(* PLC project Gaia V7.project, CODESYS CODESYS V3.5 SP22 Patch 2 *)
(* stored: creationDateTime 2026-11-05T09:22:17.1049023, modificationDateTime 2026-11-05T09:04:31.1849933 *)

TYPE DUT_COM_ADM100W : STRUCT
  COM_INPUT_IR : ARRAY[0..87] OF WORD;  (* [COM : Modbus RTU, input (equipment to PLC)] Input registers 0..87, 32-bit float, MSW first (ABCD) *)
  COM_INPUT_COILS : ARRAY[0..1] OF BYTE;  (* Coils 0..9 = alarms 1..10 (byte.bit) *)
  HMI_INPUT_LOCAL_REQUEST : BOOL;  (* [HMI (local PanelView) : input (to PLC)] Coil 12 | ADM100W Local Request *)
  HMI_INPUT_AUTO_REQUEST : BOOL;  (* Coil 13 | ADM100W Auto Request *)
  HMI_OUTPUT_ALARM_1_STATUS : BOOL;  (* [HMI (local PanelView) : output (from PLC)] DI 10003 | ADM100W Alarm 1 Status *)
  HMI_OUTPUT_ALARM_2_STATUS : BOOL;  (* DI 10004 | ADM100W Alarm 2 Status *)
  HMI_OUTPUT_ALARM_3_STATUS : BOOL;  (* DI 10005 | ADM100W Alarm 3 Status *)
  HMI_OUTPUT_ALARM_4_STATUS : BOOL;  (* DI 10006 | ADM100W Alarm 4 Status *)
  HMI_OUTPUT_ALARM_5_STATUS : BOOL;  (* DI 10007 | ADM100W Alarm 5 Status *)
  HMI_OUTPUT_ALARM_6_STATUS : BOOL;  (* DI 10008 | ADM100W Alarm 6 Status *)
  HMI_OUTPUT_ALARM_7_STATUS : BOOL;  (* DI 10009 | ADM100W Alarm 7 Status *)
  HMI_OUTPUT_ALARM_8_STATUS : BOOL;  (* DI 10010 | ADM100W Alarm 8 Status *)
  HMI_OUTPUT_ALARM_9_STATUS : BOOL;  (* DI 10011 | ADM100W Alarm 9 Status *)
  HMI_OUTPUT_ALARM_10_STATUS : BOOL;  (* DI 10012 | ADM100W Alarm 10 Status *)
  HMI_OUTPUT_LOCAL_ACTIVE : BOOL;  (* DI 10018 | ADM100W Local Active *)
  HMI_OUTPUT_FREQUENCY : DUT_Union_Real_Word;  (* IR 1-2 | ADM100W Frequency | Hz *)
  HMI_OUTPUT_L1_L2_VOLTAGE : DUT_Union_Real_Word;  (* IR 3-4 | ADM100W L1-L2 Voltage | V *)
  HMI_OUTPUT_L1_N_VOLTAGE : DUT_Union_Real_Word;  (* IR 5-6 | ADM100W L1-N Voltage | V *)
  HMI_OUTPUT_L1_CURRENT : DUT_Union_Real_Word;  (* IR 7-8 | ADM100W L1 Current | A *)
  HMI_OUTPUT_L1_ACTIVE_POWER : DUT_Union_Real_Word;  (* IR 9-10 | ADM100W L1 Active Power *)
  HMI_OUTPUT_L1_APPARENT_POWER : DUT_Union_Real_Word;  (* IR 11-12 | ADM100W L1 Apparent Power *)
  HMI_OUTPUT_L1_REACTIVE_POWER : DUT_Union_Real_Word;  (* IR 13-14 | ADM100W L1 Reactive Power *)
  HMI_OUTPUT_L1_CURRENT_PHASE_ANGLE : DUT_Union_Real_Word;  (* IR 15-16 | ADM100W L1 Current Phase Angle | deg *)
  HMI_OUTPUT_L1_POWER_FACTOR : DUT_Union_Real_Word;  (* IR 17-18 | ADM100W L1 Power Factor *)
  HMI_OUTPUT_L1_VOLTAGE_THD : DUT_Union_Real_Word;  (* IR 19-20 | ADM100W L1 Voltage THD | % *)
  HMI_OUTPUT_L1_CURRENT_THD : DUT_Union_Real_Word;  (* IR 21-22 | ADM100W L1 Current THD | % *)
  HMI_OUTPUT_L1_MAX_LOAD : DUT_Union_Real_Word;  (* IR 23-24 | ADM100W L1 Max Load *)
  HMI_OUTPUT_L1_L2_VOLTAGE_PHASE_ANGLE : DUT_Union_Real_Word;  (* IR 25-26 | ADM100W L1-L2 Voltage Phase Angle | deg *)
  HMI_OUTPUT_L2_L3_VOLTAGE : DUT_Union_Real_Word;  (* IR 27-28 | ADM100W L2-L3 Voltage | V *)
  HMI_OUTPUT_L2_N_VOLTAGE : DUT_Union_Real_Word;  (* IR 29-30 | ADM100W L2-N Voltage | V *)
  HMI_OUTPUT_L2_CURRENT : DUT_Union_Real_Word;  (* IR 31-32 | ADM100W L2 Current | A *)
  HMI_OUTPUT_L2_ACTIVE_POWER : DUT_Union_Real_Word;  (* IR 33-34 | ADM100W L2 Active Power *)
  HMI_OUTPUT_L2_APPARENT_POWER : DUT_Union_Real_Word;  (* IR 35-36 | ADM100W L2 Apparent Power *)
  HMI_OUTPUT_L2_REACTIVE_POWER : DUT_Union_Real_Word;  (* IR 37-38 | ADM100W L2 Reactive Power *)
  HMI_OUTPUT_L2_CURRENT_PHASE_ANGLE : DUT_Union_Real_Word;  (* IR 39-40 | ADM100W L2 Current Phase Angle | deg *)
  HMI_OUTPUT_L2_POWER_FACTOR : DUT_Union_Real_Word;  (* IR 41-42 | ADM100W L2 Power Factor *)
  HMI_OUTPUT_L2_VOLTAGE_THD : DUT_Union_Real_Word;  (* IR 43-44 | ADM100W L2 Voltage THD | % *)
  HMI_OUTPUT_L2_CURRENT_THD : DUT_Union_Real_Word;  (* IR 45-46 | ADM100W L2 Current THD | % *)
  HMI_OUTPUT_L2_MAX_LOAD : DUT_Union_Real_Word;  (* IR 47-48 | ADM100W L2 Max Load *)
  HMI_OUTPUT_L1_L3_VOLTAGE_PHASE_ANGLE : DUT_Union_Real_Word;  (* IR 49-50 | ADM100W L1-L3 Voltage Phase Angle | deg *)
  HMI_OUTPUT_L3_L1_VOLTAGE : DUT_Union_Real_Word;  (* IR 51-52 | ADM100W L3-L1 Voltage | V *)
  HMI_OUTPUT_L3_N_VOLTAGE : DUT_Union_Real_Word;  (* IR 53-54 | ADM100W L3-N Voltage | V *)
  HMI_OUTPUT_L3_CURRENT : DUT_Union_Real_Word;  (* IR 55-56 | ADM100W L3 Current | A *)
  HMI_OUTPUT_L3_ACTIVE_POWER : DUT_Union_Real_Word;  (* IR 57-58 | ADM100W L3 Active Power *)
  HMI_OUTPUT_L3_APPARENT_POWER : DUT_Union_Real_Word;  (* IR 59-60 | ADM100W L3 Apparent Power *)
  HMI_OUTPUT_L3_REACTIVE_POWER : DUT_Union_Real_Word;  (* IR 61-62 | ADM100W L3 Reactive Power *)
  HMI_OUTPUT_L3_CURRENT_PHASE_ANGLE : DUT_Union_Real_Word;  (* IR 63-64 | ADM100W L3 Current Phase Angle | deg *)
  HMI_OUTPUT_L3_POWER_FACTOR : DUT_Union_Real_Word;  (* IR 65-66 | ADM100W L3 Power Factor *)
  HMI_OUTPUT_L3_VOLTAGE_THD : DUT_Union_Real_Word;  (* IR 67-68 | ADM100W L3 Voltage THD | % *)
  HMI_OUTPUT_L3_CURRENT_THD : DUT_Union_Real_Word;  (* IR 69-70 | ADM100W L3 Current THD | % *)
  HMI_OUTPUT_L3_MAX_LOAD : DUT_Union_Real_Word;  (* IR 71-72 | ADM100W L3 Max Load *)
  HMI_OUTPUT_INTERNAL_TEMPERATURE : DUT_Union_Real_Word;  (* IR 73-74 | ADM100W Internal Temperature *)
  HMI_OUTPUT_ACTIVE_ENERGY : DUT_Union_Real_Word;  (* IR 75-76 | ADM100W Active Energy *)
  HMI_OUTPUT_APPARENT_ENERGY : DUT_Union_Real_Word;  (* IR 77-78 | ADM100W Apparent Energy *)
  HMI_OUTPUT_REACTIVE_ENERGY : DUT_Union_Real_Word;  (* IR 79-80 | ADM100W Reactive Energy *)
  HMI_OUTPUT_TOTAL_ACTIVE_POWER : DUT_Union_Real_Word;  (* IR 81-82 | ADM100W Total Active Power *)
  HMI_OUTPUT_TOTAL_APPARENT_POWER : DUT_Union_Real_Word;  (* IR 83-84 | ADM100W Total Apparent Power *)
  HMI_OUTPUT_TOTAL_REACTIVE_POWER : DUT_Union_Real_Word;  (* IR 85-86 | ADM100W Total Reactive Power *)
  HMI_OUTPUT_ALL_PHASE_POWER_FACTOR : DUT_Union_Real_Word;  (* IR 87-88 | ADM100W All Phase Power Factor *)
END_STRUCT;
END_TYPE

TYPE DUT_COM_DIP1500 : STRUCT
  COM_INPUT_IR : ARRAY[0..4] OF WORD;  (* [COM : Modbus RTU, input (equipment to PLC)] Input registers 0x3001..0x3005 *)
  COM_INPUT_HR_COUNTERS : ARRAY[0..3] OF WORD;  (* Holding registers 0x4007..0x400A (read) *)
  COM_OUTPUT_COILS : ARRAY[0..3] OF BOOL;  (* [COM : Modbus RTU, output (PLC to equipment)] Coils 0x0001..0x0004 *)
  COM_OUTPUT_HR_CMD : ARRAY[0..5] OF WORD;  (* Holding registers 0x4001..0x4006 (write) *)
  COM_OUTPUT_HR_CONFIG : ARRAY[0..6] OF WORD;  (* Holding registers 0x400B..0x4011 (write) *)
  COM_OUTPUT_CMD_TRIGGER : BOOL;  (* Rising edge trigger of the command write channel(s), mapped in the Modbus slave I/O mapping *)
  COM_OUTPUT_CONFIG_TRIGGER : BOOL;  (* Rising edge trigger of the configuration write channel, mapped in the Modbus slave I/O mapping *)
  HMI_INPUT_MOTOR_START_STOP : BOOL;  (* [HMI (local PanelView) : input (to PLC)] Coil 3 | DIP1500 Motor Start Stop *)
  HMI_INPUT_MOTOR_DIRECTION : BOOL;  (* Coil 4 | DIP1500 Motor Direction *)
  HMI_INPUT_FLASH_SAVE : BOOL;  (* Coil 5 | DIP1500 Flash Save *)
  HMI_INPUT_OPERATION_MODE : BOOL;  (* Coil 6 | DIP1500 Operation Mode *)
  HMI_INPUT_PARAM_WRITE_ENABLE : BOOL;  (* Coil 7 | DIP1500 Parameter Write Enable *)
  HMI_INPUT_LOCAL_REQUEST : BOOL;  (* Coil 10 | DIP1500 Local Request *)
  HMI_INPUT_AUTO_REQUEST : BOOL;  (* Coil 11 | DIP1500 Auto Request *)
  HMI_INPUT_FOOT_SWITCH_INPUT_MODE : WORD;  (* HR 9 | DIP1500 Foot Switch Input Mode *)
  HMI_INPUT_LIQUID_LEVEL_INPUT_MODE : WORD;  (* HR 10 | DIP1500 Liquid Level Input Mode *)
  HMI_INPUT_STATE_OUTPUT_MODE : WORD;  (* HR 11 | DIP1500 State Output Mode *)
  HMI_INPUT_COMMUNICATION_ADDRESS : WORD;  (* HR 12 | DIP1500 Communication Address *)
  HMI_INPUT_BAUD_RATE_INDEX : WORD;  (* HR 13 | DIP1500 Baud Rate Index | index *)
  HMI_INPUT_MOTOR_SPEED : DUT_Union_Real_Word;  (* HR 1-2 | DIP1500 Motor Speed | rpm *)
  HMI_INPUT_MAX_MOTOR_SPEED : DUT_Union_Real_Word;  (* HR 3-4 | DIP1500 Max Motor Speed | rpm *)
  HMI_INPUT_RUN_TIME_OR_VOLUME_SETPOINT : DUT_Union_Real_Word;  (* HR 5-6 | DIP1500 Run Time Or Volume Setpoint | ms (time mode) / ml (volume mode) *)
  HMI_INPUT_FLOW_RATE_OR_SPEED_CALIBRATION_COEFFICIENT : DUT_Union_Real_Word;  (* HR 7-8 | DIP1500 Flow Rate Or Speed Calibration Coefficient | ml/min or rpm *)
  HMI_OUTPUT_LOCAL_ACTIVE : BOOL;  (* [HMI (local PanelView) : output (from PLC)] DI 10016 | DIP1500 Local Active *)
  HMI_OUTPUT_FIRMWARE_VERSION : WORD;  (* IR 91 | DIP1500 Firmware Version | 3+5+8 bits (major+minor+revision) *)
  HMI_OUTPUT_HARDWARE_VERSION : WORD;  (* IR 92 | DIP1500 Hardware Version | 3+5+8 bits (major+minor+revision) *)
  HMI_OUTPUT_TEMPERATURE : WORD;  (* IR 93 | DIP1500 Temperature | degC | (raw - 500) / 10 *)
  HMI_OUTPUT_FLOAT_LEVEL_ALARM : WORD;  (* IR 94 | DIP1500 Float Level Alarm *)
  HMI_OUTPUT_DIGITAL_OUTPUT_VALUE : WORD;  (* IR 95 | DIP1500 Digital Output Value *)
  HMI_OUTPUT_REAL_TIME_RUN_TIME_OR_VOLUME : DUT_Union_Real_Word;  (* IR 96-97 | DIP1500 Real-Time Run Time Or Volume | ms (time mode) / ml (volume mode) *)
  HMI_OUTPUT_ACCUMULATED_RUN_TIME_OR_VOLUME : DUT_Union_Real_Word;  (* IR 98-99 | DIP1500 Accumulated Run Time Or Volume | ms (time mode) / ml (volume mode) *)
END_STRUCT;
END_TYPE

TYPE DUT_COM_DOSENSOR : STRUCT
  HMI_INPUT_CALIBRATION_HIGH : BOOL;  (* [HMI (local PanelView) : input (to PLC)] Coil 1 | DO Calibration High *)
  HMI_INPUT_CALIBRATION_LOW : BOOL;  (* Coil 2 | DO Calibration Low *)
  HMI_INPUT_LOCAL_REQUEST : BOOL;  (* Coil 8 | DO Sensor Local Request *)
  HMI_INPUT_AUTO_REQUEST : BOOL;  (* Coil 9 | DO Sensor Auto Request *)
  HMI_OUTPUT_FAULT : BOOL;  (* [HMI (local PanelView) : output (from PLC)] DI 10001 | Do sensor fault *)
  HMI_OUTPUT_CALIBRATION_DONE : BOOL;  (* DI 10002 | Do sensor calibration done *)
  HMI_OUTPUT_LOCAL_ACTIVE : BOOL;  (* DI 10014 | DO Sensor Local Active *)
  HMI_OUTPUT_SIGNAL : DUT_Union_Real_Word;  (* IR 89-90 | DO Sensor Signal *)
END_STRUCT;
END_TYPE

TYPE DUT_COM_UPI_LOCAL_HMI : STRUCT
  HMI_INPUT_LOCAL_REQUEST : BOOL;  (* [HMI (local PanelView) : input (to PLC)] Coil 14 | Global Local HMI Request *)
  HMI_INPUT_AUTO_REQUEST : BOOL;  (* Coil 15 | Global Auto HMI Request *)
  HMI_OUTPUT_LOCAL_ACTIVE : BOOL;  (* [HMI (local PanelView) : output (from PLC)] DI 10020 | Global Local HMI Active *)
END_STRUCT;
END_TYPE

TYPE DUT_EXC_ADM100W : STRUCT
  EXC_OUTPUT_FREQUENCY : REAL;  (* [EXC : to other equipment] Hz *)
  EXC_OUTPUT_L1_N_VOLTAGE : REAL;  (* V *)
  EXC_OUTPUT_L1_CURRENT : REAL;  (* A *)
  EXC_OUTPUT_L1_ACTIVE_POWER : REAL;  (* W *)
  EXC_OUTPUT_L1_APPARENT_POWER : REAL;  (* VA *)
  EXC_OUTPUT_L1_REACTIVE_POWER : REAL;  (* VAr *)
  EXC_OUTPUT_L1_POWER_FACTOR : REAL;  (* - *)
  EXC_OUTPUT_L1_VOLTAGE_THD : REAL;  (* % *)
  EXC_OUTPUT_L1_CURRENT_THD : REAL;  (* % *)
  EXC_OUTPUT_L1_MAX_LOAD : REAL;  (* % of 60 A *)
  EXC_OUTPUT_INTERNAL_TEMPERATURE : REAL;  (* degC *)
  EXC_OUTPUT_ACTIVE_ENERGY : REAL;  (* kWh *)
  EXC_OUTPUT_DATA_VALID : BOOL;  (* FALSE = values not usable. Not managed yet (no Modbus diagnostic) *)
  UPI_INPUT_GLOBAL_LOCAL_HMI : BOOL;  (* [UPI : functional units to equipment] From UPI_LOCAL_HMI : global HMI local active *)
END_STRUCT;
END_TYPE

TYPE DUT_EXC_DIP1500 : STRUCT
  UPI_INPUT_GLOBAL_LOCAL_HMI : BOOL;  (* [UPI : functional units to equipment] From UPI_LOCAL_HMI : global HMI local active *)
  UPI_INPUT_RUN : BOOL;  (* [UPI : commands used in auto mode] Auto mode command : run *)
  UPI_INPUT_CLOCKWISE : BOOL;  (* Auto mode command : 1 clockwise *)
  UPI_INPUT_VOLUME_MODE : BOOL;  (* Auto mode command : 0 time mode, 1 volume mode *)
  UPI_INPUT_SPEED : REAL;  (* Auto mode command : speed, rpm *)
  UPI_INPUT_RUN_SETPOINT : REAL;  (* Auto mode command : ms (time mode) or ml (volume mode), 0 = continuous *)
END_STRUCT;
END_TYPE

TYPE DUT_EXC_DOSENSOR : STRUCT
  EXC_OUTPUT_SIGNAL : REAL;  (* [EXC : to other equipment] Dissolved oxygen measure *)
  UPI_INPUT_GLOBAL_LOCAL_HMI : BOOL;  (* [UPI : functional units to equipment] From UPI_LOCAL_HMI : global HMI local active *)
END_STRUCT;
END_TYPE

TYPE DUT_EXC_UPI_LOCAL_HMI : STRUCT
  UPI_OUTPUT_LOCAL_ACTIVE : BOOL;  (* [UPI : to equipment] Global HMI local active *)
END_STRUCT;
END_TYPE

TYPE DUT_INT_ADM100W : STRUCT
  HMI_LOCAL_REQUEST : BOOL;  (* [Control mode] From HMI : local request (pulse or maintained) *)
  HMI_AUTO_REQUEST : BOOL;  (* From HMI : auto request, releases the individual HMI local *)
  GLOBAL_LOCAL_HMI : BOOL;  (* From UPI_LOCAL_HMI : global HMI local active *)
  LOCAL_HMI_INDIVIDUAL : BOOL;  (* Memory : individual HMI local, set by local request, reset by auto request *)
  LOCAL_HMI : BOOL;  (* Result : equipment in HMI local (individual or global) *)
  AUTO : BOOL;  (* Result : no local mode, commands come from the functional units (UPI) *)
  ALARM_1 : BOOL;  (* [Alarms] Alarm 1 status *)
  ALARM_2 : BOOL;  (* Alarm 2 status *)
  ALARM_3 : BOOL;  (* Alarm 3 status *)
  ALARM_4 : BOOL;  (* Alarm 4 status *)
  ALARM_5 : BOOL;  (* Alarm 5 status *)
  ALARM_6 : BOOL;  (* Alarm 6 status *)
  ALARM_7 : BOOL;  (* Alarm 7 status *)
  ALARM_8 : BOOL;  (* Alarm 8 status *)
  ALARM_9 : BOOL;  (* Alarm 9 status *)
  ALARM_10 : BOOL;  (* Alarm 10 status *)
  FREQUENCY : REAL;  (* [Measures] Frequency | Hz *)
  L1_L2_VOLTAGE : REAL;  (* L1-L2 Voltage | V *)
  L1_N_VOLTAGE : REAL;  (* L1-N Voltage | V *)
  L1_CURRENT : REAL;  (* L1 Current | A *)
  L1_ACTIVE_POWER : REAL;  (* L1 Active Power | W *)
  L1_APPARENT_POWER : REAL;  (* L1 Apparent Power | VA *)
  L1_REACTIVE_POWER : REAL;  (* L1 Reactive Power | W *)
  L1_CURRENT_PHASE_ANGLE : REAL;  (* L1 Current Phase Angle | deg *)
  L1_POWER_FACTOR : REAL;  (* L1 Power Factor | - *)
  L1_VOLTAGE_THD : REAL;  (* L1 Voltage THD | % *)
  L1_CURRENT_THD : REAL;  (* L1 Current THD | % *)
  L1_MAX_LOAD : REAL;  (* L1 Max Load | % of 60 A *)
  L1_L2_VOLTAGE_PHASE_ANGLE : REAL;  (* L1-L2 Voltage Phase Angle | deg *)
  L2_L3_VOLTAGE : REAL;  (* L2-L3 Voltage | V *)
  L2_N_VOLTAGE : REAL;  (* L2-N Voltage | V *)
  L2_CURRENT : REAL;  (* L2 Current | A *)
  L2_ACTIVE_POWER : REAL;  (* L2 Active Power | W *)
  L2_APPARENT_POWER : REAL;  (* L2 Apparent Power | VA *)
  L2_REACTIVE_POWER : REAL;  (* L2 Reactive Power | W *)
  L2_CURRENT_PHASE_ANGLE : REAL;  (* L2 Current Phase Angle | deg *)
  L2_POWER_FACTOR : REAL;  (* L2 Power Factor | - *)
  L2_VOLTAGE_THD : REAL;  (* L2 Voltage THD | % *)
  L2_CURRENT_THD : REAL;  (* L2 Current THD | % *)
  L2_MAX_LOAD : REAL;  (* L2 Max Load | % of 60 A *)
  L1_L3_VOLTAGE_PHASE_ANGLE : REAL;  (* L1-L3 Voltage Phase Angle | deg *)
  L3_L1_VOLTAGE : REAL;  (* L3-L1 Voltage | V *)
  L3_N_VOLTAGE : REAL;  (* L3-N Voltage | V *)
  L3_CURRENT : REAL;  (* L3 Current | A *)
  L3_ACTIVE_POWER : REAL;  (* L3 Active Power | W *)
  L3_APPARENT_POWER : REAL;  (* L3 Apparent Power | VA *)
  L3_REACTIVE_POWER : REAL;  (* L3 Reactive Power | W *)
  L3_CURRENT_PHASE_ANGLE : REAL;  (* L3 Current Phase Angle | deg *)
  L3_POWER_FACTOR : REAL;  (* L3 Power Factor | - *)
  L3_VOLTAGE_THD : REAL;  (* L3 Voltage THD | % *)
  L3_CURRENT_THD : REAL;  (* L3 Current THD | % *)
  L3_MAX_LOAD : REAL;  (* L3 Max Load | % of 60 A *)
  INTERNAL_TEMPERATURE : REAL;  (* Internal Temperature | degC *)
  ACTIVE_ENERGY : REAL;  (* Active Energy | kWh *)
  APPARENT_ENERGY : REAL;  (* Apparent Energy | per ADM100W config *)
  REACTIVE_ENERGY : REAL;  (* Reactive Energy | kWh *)
  TOTAL_ACTIVE_POWER : REAL;  (* Total Active Power | W *)
  TOTAL_APPARENT_POWER : REAL;  (* Total Apparent Power | VA *)
  TOTAL_REACTIVE_POWER : REAL;  (* Total Reactive Power | W *)
  ALL_PHASE_POWER_FACTOR : REAL;  (* All Phase Power Factor | - *)
END_STRUCT;
END_TYPE

TYPE DUT_INT_DIP1500 : STRUCT
  HMI_LOCAL_REQUEST : BOOL;  (* [Control mode] From HMI : local request (pulse or maintained) *)
  HMI_AUTO_REQUEST : BOOL;  (* From HMI : auto request, releases the individual HMI local *)
  GLOBAL_LOCAL_HMI : BOOL;  (* From UPI_LOCAL_HMI : global HMI local active *)
  LOCAL_HMI_INDIVIDUAL : BOOL;  (* Memory : individual HMI local, set by local request, reset by auto request *)
  LOCAL_HMI : BOOL;  (* Result : equipment in HMI local (individual or global) *)
  AUTO : BOOL;  (* Result : no local mode, commands come from the functional units (UPI) *)
  CMD_RUN : BOOL;  (* [Commands (to pump), from the active source] 0 stop, 1 start *)
  CMD_CLOCKWISE : BOOL;  (* 0 counterclockwise, 1 clockwise *)
  CMD_SAVE_FLASH : BOOL;  (* 1 s pulse to coil 0x0003, saves pump parameters to flash *)
  CMD_VOLUME_MODE : BOOL;  (* 0 time mode, 1 volume mode *)
  CMD_SPEED : REAL;  (* rpm *)
  CMD_MAX_SPEED : REAL;  (* rpm *)
  CMD_RUN_SETPOINT : REAL;  (* ms (time mode) or ml (volume mode), 0 = continuous *)
  CMD_CALIB_COEF : REAL;  (* ml/min or rpm *)
  CMD_FOOT_MODE : WORD;  (* Foot switch input mode *)
  CMD_LEVEL_MODE : WORD;  (* Liquid level input mode *)
  CMD_STATE_OUT_MODE : WORD;  (* State output mode *)
  CMD_ADDRESS : WORD;  (* Modbus address *)
  CMD_BAUD_INDEX : WORD;  (* 0=1200 .. 3=9600 .. 7=115200 *)
  PARAM_WRITE_ENABLE : BOOL;  (* [Parameter writing] 1 = write configuration to the pump, 0 = stop writing *)
  FLASH_SAVE_REQUEST : BOOL;  (* Flash save request (rising edge used) *)
  PARAM_VALID : BOOL;  (* Address 1..31, baud index 0..7, max speed > 0, calibration coefficient > 0 *)
  PULSE_500MS : BOOL;  (* [Write triggers] Square wave, 500 ms period, source of the trigger edges *)
  CMD_CHANGED : BOOL;  (* A command value changed this cycle *)
  CMD_WINDOW : BOOL;  (* Command write window, 3 s after the last change *)
  CMD_TRIGGER : BOOL;  (* Command channel trigger *)
  CONFIG_TRIGGER : BOOL;  (* Configuration channel trigger *)
  PREV_RUN : BOOL;  (* [Previous command values] Previous values for change detection *)
  PREV_CLOCKWISE : BOOL;
  PREV_VOLUME_MODE : BOOL;
  PREV_SAVE_FLASH : BOOL;
  PREV_SPEED : REAL;
  PREV_MAX_SPEED : REAL;
  PREV_RUN_SETPOINT : REAL;
  FBK_FIRMWARE_VERSION : WORD;  (* [Feedback (from pump)] 3+5+8 bits (major+minor+revision) *)
  FBK_HARDWARE_VERSION : WORD;  (* 3+5+8 bits (major+sub+reserved) *)
  FBK_TEMPERATURE : WORD;  (* (raw - 500) / 10 = degC, 65535 = not connected *)
  FBK_LEVEL_ALARM : WORD;  (* 0 no alarm, 1 alarm, 65535 = not connected *)
  FBK_DIGITAL_OUTPUT : WORD;  (* Digital output value *)
  FBK_RUN_ACTUAL : REAL;  (* Current run, ms (time mode) or ml (volume mode) *)
  FBK_RUN_TOTAL : REAL;  (* Accumulated run, ms (time mode) or ml (volume mode) *)
  UDINT_TEMP : UDINT;  (* [Work] Work variable, time mode conversion *)
  SRC_MAX_MOTOR_SPEED : REAL;  (* [Parameter source] Value typed in the active local supervision *)
  SRC_CALIBRATION_COEFFICIENT : REAL;
  SRC_FOOT_SWITCH_INPUT_MODE : WORD;
  SRC_LIQUID_LEVEL_INPUT_MODE : WORD;
  SRC_STATE_OUTPUT_MODE : WORD;
  SRC_COMMUNICATION_ADDRESS : WORD;
  SRC_BAUD_RATE_INDEX : WORD;
  PREV_SRC_MAX_MOTOR_SPEED : REAL;  (* [Parameter change detection] Previous source values *)
  PREV_SRC_CALIBRATION_COEFFICIENT : REAL;
  PREV_SRC_FOOT_SWITCH_INPUT_MODE : WORD;
  PREV_SRC_LIQUID_LEVEL_INPUT_MODE : WORD;
  PREV_SRC_STATE_OUTPUT_MODE : WORD;
  PREV_SRC_COMMUNICATION_ADDRESS : WORD;
  PREV_SRC_BAUD_RATE_INDEX : WORD;
  PREV_LOCAL_HMI : BOOL;
  SOURCE_CHANGED : BOOL;  (* The active local source changed this cycle : no parameter is taken *)
END_STRUCT;
END_TYPE

TYPE DUT_INT_DOSENSOR : STRUCT
  HMI_LOCAL_REQUEST : BOOL;  (* [Control mode] From HMI : local request (pulse or maintained) *)
  HMI_AUTO_REQUEST : BOOL;  (* From HMI : auto request, releases the individual HMI local *)
  GLOBAL_LOCAL_HMI : BOOL;  (* From UPI_LOCAL_HMI : global HMI local active *)
  LOCAL_HMI_INDIVIDUAL : BOOL;  (* Memory : individual HMI local, set by local request, reset by auto request *)
  LOCAL_HMI : BOOL;  (* Result : equipment in HMI local (individual or global) *)
  AUTO : BOOL;  (* Result : no local mode, commands come from the functional units (UPI) *)
  SIGNAL_RAW : DWORD;  (* [Inputs] Raw analog input *)
  FAULT : BOOL;  (* Sensor fault (digital input) *)
  CALIB_HIGH_REQUEST : BOOL;  (* High calibration request from the active source *)
  CALIB_LOW_REQUEST : BOOL;  (* Low calibration request from the active source *)
  SIGNAL : REAL;  (* [Results] Scaled measure *)
  CALIB_HIGH : BOOL;  (* High calibration pulse to sensor (1 s) *)
  CALIB_LOW : BOOL;  (* Low calibration pulse to sensor (1 s) *)
  CALIB_DONE : BOOL;  (* Calibration done message (5 s) *)
END_STRUCT;
END_TYPE

TYPE DUT_INT_UPI_LOCAL_HMI : STRUCT
  LOCAL_REQUEST : BOOL;  (* Local request (pulse or maintained) *)
  AUTO_REQUEST : BOOL;  (* Auto request, releases the global local *)
  LOCAL_ACTIVE : BOOL;  (* Memory : global local active *)
END_STRUCT;
END_TYPE

TYPE DUT_IO_ADM100W : STRUCT
  SPARE : BOOL;  (* Placeholder, structure not used yet *)
END_STRUCT;
END_TYPE

TYPE DUT_IO_DIP1500 : STRUCT
  SPARE : BOOL;  (* Placeholder, structure not used yet *)
END_STRUCT;
END_TYPE

TYPE DUT_IO_DOSENSOR : STRUCT
  INPUT_SIGNAL : DWORD;  (* [INPUT (field to PLC)] Analog input, raw value *)
  INPUT_SENSOR_FAULT : BOOL;  (* Digital input, sensor fault *)
  OUTPUT_CALIBRATION_HIGH : BOOL;  (* [OUTPUT (PLC to field)] Digital output, high calibration *)
  OUTPUT_CALIBRATION_LOW : BOOL;  (* Digital output, low calibration *)
END_STRUCT;
END_TYPE

TYPE DUT_PA_ADM100W : STRUCT
  SPARE : BOOL;  (* Placeholder, structure not used yet *)
END_STRUCT;
END_TYPE

TYPE DUT_PA_DIP1500 : STRUCT
  MAX_MOTOR_SPEED : REAL := 350;  (* [Pump configuration, default value = declaration value, kept in GVL_PA (persistent)] rpm. Max motor speed (pump register 0x4003) *)
  CALIBRATION_COEFFICIENT : REAL := 100;  (* ml/min or rpm. Flow / speed calibration coefficient (0x400B) *)
  FOOT_SWITCH_INPUT_MODE : WORD := 0;  (* Foot switch input mode (0x400D) *)
  LIQUID_LEVEL_INPUT_MODE : WORD := 100;  (* Liquid level input mode (0x400E) *)
  STATE_OUTPUT_MODE : WORD := 7;  (* State output mode (0x400F) *)
  COMMUNICATION_ADDRESS : WORD := 11;  (* Pump Modbus address, 1..31 (0x4010) *)
  BAUD_RATE_INDEX : WORD := 3;  (* 0=1200 .. 3=9600 .. 7=115200 (0x4011) *)
END_STRUCT;
END_TYPE

TYPE DUT_PA_DOSENSOR : STRUCT
  SPARE : BOOL;  (* Placeholder, structure not used yet *)
END_STRUCT;
END_TYPE

TYPE DUT_Union_Real_Word : UNION
  Real_value : REAL;
  Word_value : ARRAY[0..1] OF WORD;
END_UNION;
END_TYPE

FUNCTION_BLOCK FB_INST_ADM100W
  VAR_IN_OUT
    PA : DUT_PA_ADM100W;  (* Parameters (persistent, GVL_PA) *)
    COM : DUT_COM_ADM100W;  (* Communication : Modbus RTU (COM_), HMI PanelView (HMI_) *)
    EXC : DUT_EXC_ADM100W;  (* Exchanges : other equipment (EXC_), functional units (UPI_) *)
    IO : DUT_IO_ADM100W;  (* Wired PLC I/O *)
  END_VAR
  VAR
    INTERN : DUT_INT_ADM100W;  (* Internal variables *)
  END_VAR

                  
//==============================================================================
// FB_INST_ADM100W
// Trumeter ADM100W power meter, Modbus RTU, 32-bit float MSW first (ABCD). No command : local mode is only reported
// 1. INPUTS     : requests, control mode, command source, equipment feedback -> INTERN
// 2. PROCESSING : on INTERN only
// 3. OUTPUTS    : INTERN -> COM / IO / EXC
// Control mode  : local HMI (individual or global) > auto (functional units)
//==============================================================================

//------------------------------------------------------------------------------
// 1. INPUTS
//------------------------------------------------------------------------------
	//--- Control mode requests (HMI, global HMI local from UPI_LOCAL_HMI)
	INTERN.HMI_LOCAL_REQUEST := COM.HMI_INPUT_LOCAL_REQUEST;
	INTERN.HMI_AUTO_REQUEST  := COM.HMI_INPUT_AUTO_REQUEST;
	INTERN.GLOBAL_LOCAL_HMI  := EXC.UPI_INPUT_GLOBAL_LOCAL_HMI;

	//--- Control mode
	// Individual memory : set by the local request, reset by the auto request (auto wins if both)
	IF INTERN.HMI_LOCAL_REQUEST THEN
		INTERN.LOCAL_HMI_INDIVIDUAL := TRUE;
	END_IF
	IF INTERN.HMI_AUTO_REQUEST THEN
		INTERN.LOCAL_HMI_INDIVIDUAL := FALSE;
	END_IF

	// Resulting mode : HMI local (individual OR global), otherwise auto
	INTERN.LOCAL_HMI := INTERN.LOCAL_HMI_INDIVIDUAL OR INTERN.GLOBAL_LOCAL_HMI;
	INTERN.AUTO      := NOT INTERN.LOCAL_HMI;

	//--- COM : alarms (coils 0..9)
	INTERN.ALARM_1  := COM.COM_INPUT_COILS[0].0;
	INTERN.ALARM_2  := COM.COM_INPUT_COILS[0].1;
	INTERN.ALARM_3  := COM.COM_INPUT_COILS[0].2;
	INTERN.ALARM_4  := COM.COM_INPUT_COILS[0].3;
	INTERN.ALARM_5  := COM.COM_INPUT_COILS[0].4;
	INTERN.ALARM_6  := COM.COM_INPUT_COILS[0].5;
	INTERN.ALARM_7  := COM.COM_INPUT_COILS[0].6;
	INTERN.ALARM_8  := COM.COM_INPUT_COILS[0].7;
	INTERN.ALARM_9  := COM.COM_INPUT_COILS[1].0;
	INTERN.ALARM_10 := COM.COM_INPUT_COILS[1].1;

	//--- COM : measures (input registers, MSW first)
	INTERN.FREQUENCY                 := FNC_WORDS_TO_REAL(High_word := COM.COM_INPUT_IR[0], Low_word := COM.COM_INPUT_IR[1]);
	INTERN.L1_L2_VOLTAGE             := FNC_WORDS_TO_REAL(High_word := COM.COM_INPUT_IR[2], Low_word := COM.COM_INPUT_IR[3]);
	INTERN.L1_N_VOLTAGE              := FNC_WORDS_TO_REAL(High_word := COM.COM_INPUT_IR[4], Low_word := COM.COM_INPUT_IR[5]);
	INTERN.L1_CURRENT                := FNC_WORDS_TO_REAL(High_word := COM.COM_INPUT_IR[6], Low_word := COM.COM_INPUT_IR[7]);
	INTERN.L1_ACTIVE_POWER           := FNC_WORDS_TO_REAL(High_word := COM.COM_INPUT_IR[8], Low_word := COM.COM_INPUT_IR[9]);
	INTERN.L1_APPARENT_POWER         := FNC_WORDS_TO_REAL(High_word := COM.COM_INPUT_IR[10], Low_word := COM.COM_INPUT_IR[11]);
	INTERN.L1_REACTIVE_POWER         := FNC_WORDS_TO_REAL(High_word := COM.COM_INPUT_IR[12], Low_word := COM.COM_INPUT_IR[13]);
	INTERN.L1_CURRENT_PHASE_ANGLE    := FNC_WORDS_TO_REAL(High_word := COM.COM_INPUT_IR[14], Low_word := COM.COM_INPUT_IR[15]);
	INTERN.L1_POWER_FACTOR           := FNC_WORDS_TO_REAL(High_word := COM.COM_INPUT_IR[16], Low_word := COM.COM_INPUT_IR[17]);
	INTERN.L1_VOLTAGE_THD            := FNC_WORDS_TO_REAL(High_word := COM.COM_INPUT_IR[18], Low_word := COM.COM_INPUT_IR[19]);
	INTERN.L1_CURRENT_THD            := FNC_WORDS_TO_REAL(High_word := COM.COM_INPUT_IR[20], Low_word := COM.COM_INPUT_IR[21]);
	INTERN.L1_MAX_LOAD               := FNC_WORDS_TO_REAL(High_word := COM.COM_INPUT_IR[22], Low_word := COM.COM_INPUT_IR[23]);
	INTERN.L1_L2_VOLTAGE_PHASE_ANGLE := FNC_WORDS_TO_REAL(High_word := COM.COM_INPUT_IR[24], Low_word := COM.COM_INPUT_IR[25]);
	INTERN.L2_L3_VOLTAGE             := FNC_WORDS_TO_REAL(High_word := COM.COM_INPUT_IR[26], Low_word := COM.COM_INPUT_IR[27]);
	INTERN.L2_N_VOLTAGE              := FNC_WORDS_TO_REAL(High_word := COM.COM_INPUT_IR[28], Low_word := COM.COM_INPUT_IR[29]);
	INTERN.L2_CURRENT                := FNC_WORDS_TO_REAL(High_word := COM.COM_INPUT_IR[30], Low_word := COM.COM_INPUT_IR[31]);
	INTERN.L2_ACTIVE_POWER           := FNC_WORDS_TO_REAL(High_word := COM.COM_INPUT_IR[32], Low_word := COM.COM_INPUT_IR[33]);
	INTERN.L2_APPARENT_POWER         := FNC_WORDS_TO_REAL(High_word := COM.COM_INPUT_IR[34], Low_word := COM.COM_INPUT_IR[35]);
	INTERN.L2_REACTIVE_POWER         := FNC_WORDS_TO_REAL(High_word := COM.COM_INPUT_IR[36], Low_word := COM.COM_INPUT_IR[37]);
	INTERN.L2_CURRENT_PHASE_ANGLE    := FNC_WORDS_TO_REAL(High_word := COM.COM_INPUT_IR[38], Low_word := COM.COM_INPUT_IR[39]);
	INTERN.L2_POWER_FACTOR           := FNC_WORDS_TO_REAL(High_word := COM.COM_INPUT_IR[40], Low_word := COM.COM_INPUT_IR[41]);
	INTERN.L2_VOLTAGE_THD            := FNC_WORDS_TO_REAL(High_word := COM.COM_INPUT_IR[42], Low_word := COM.COM_INPUT_IR[43]);
	INTERN.L2_CURRENT_THD            := FNC_WORDS_TO_REAL(High_word := COM.COM_INPUT_IR[44], Low_word := COM.COM_INPUT_IR[45]);
	INTERN.L2_MAX_LOAD               := FNC_WORDS_TO_REAL(High_word := COM.COM_INPUT_IR[46], Low_word := COM.COM_INPUT_IR[47]);
	INTERN.L1_L3_VOLTAGE_PHASE_ANGLE := FNC_WORDS_TO_REAL(High_word := COM.COM_INPUT_IR[48], Low_word := COM.COM_INPUT_IR[49]);
	INTERN.L3_L1_VOLTAGE             := FNC_WORDS_TO_REAL(High_word := COM.COM_INPUT_IR[50], Low_word := COM.COM_INPUT_IR[51]);
	INTERN.L3_N_VOLTAGE              := FNC_WORDS_TO_REAL(High_word := COM.COM_INPUT_IR[52], Low_word := COM.COM_INPUT_IR[53]);
	INTERN.L3_CURRENT                := FNC_WORDS_TO_REAL(High_word := COM.COM_INPUT_IR[54], Low_word := COM.COM_INPUT_IR[55]);
	INTERN.L3_ACTIVE_POWER           := FNC_WORDS_TO_REAL(High_word := COM.COM_INPUT_IR[56], Low_word := COM.COM_INPUT_IR[57]);
	INTERN.L3_APPARENT_POWER         := FNC_WORDS_TO_REAL(High_word := COM.COM_INPUT_IR[58], Low_word := COM.COM_INPUT_IR[59]);
	INTERN.L3_REACTIVE_POWER         := FNC_WORDS_TO_REAL(High_word := COM.COM_INPUT_IR[60], Low_word := COM.COM_INPUT_IR[61]);
	INTERN.L3_CURRENT_PHASE_ANGLE    := FNC_WORDS_TO_REAL(High_word := COM.COM_INPUT_IR[62], Low_word := COM.COM_INPUT_IR[63]);
	INTERN.L3_POWER_FACTOR           := FNC_WORDS_TO_REAL(High_word := COM.COM_INPUT_IR[64], Low_word := COM.COM_INPUT_IR[65]);
	INTERN.L3_VOLTAGE_THD            := FNC_WORDS_TO_REAL(High_word := COM.COM_INPUT_IR[66], Low_word := COM.COM_INPUT_IR[67]);
	INTERN.L3_CURRENT_THD            := FNC_WORDS_TO_REAL(High_word := COM.COM_INPUT_IR[68], Low_word := COM.COM_INPUT_IR[69]);
	INTERN.L3_MAX_LOAD               := FNC_WORDS_TO_REAL(High_word := COM.COM_INPUT_IR[70], Low_word := COM.COM_INPUT_IR[71]);
	INTERN.INTERNAL_TEMPERATURE      := FNC_WORDS_TO_REAL(High_word := COM.COM_INPUT_IR[72], Low_word := COM.COM_INPUT_IR[73]);
	INTERN.ACTIVE_ENERGY             := FNC_WORDS_TO_REAL(High_word := COM.COM_INPUT_IR[74], Low_word := COM.COM_INPUT_IR[75]);
	INTERN.APPARENT_ENERGY           := FNC_WORDS_TO_REAL(High_word := COM.COM_INPUT_IR[76], Low_word := COM.COM_INPUT_IR[77]);
	INTERN.REACTIVE_ENERGY           := FNC_WORDS_TO_REAL(High_word := COM.COM_INPUT_IR[78], Low_word := COM.COM_INPUT_IR[79]);
	INTERN.TOTAL_ACTIVE_POWER        := FNC_WORDS_TO_REAL(High_word := COM.COM_INPUT_IR[80], Low_word := COM.COM_INPUT_IR[81]);
	INTERN.TOTAL_APPARENT_POWER      := FNC_WORDS_TO_REAL(High_word := COM.COM_INPUT_IR[82], Low_word := COM.COM_INPUT_IR[83]);
	INTERN.TOTAL_REACTIVE_POWER      := FNC_WORDS_TO_REAL(High_word := COM.COM_INPUT_IR[84], Low_word := COM.COM_INPUT_IR[85]);
	INTERN.ALL_PHASE_POWER_FACTOR    := FNC_WORDS_TO_REAL(High_word := COM.COM_INPUT_IR[86], Low_word := COM.COM_INPUT_IR[87]);


//------------------------------------------------------------------------------
// 2. PROCESSING
//------------------------------------------------------------------------------
	// Nothing


//------------------------------------------------------------------------------
// 3. OUTPUTS
//------------------------------------------------------------------------------
	//--- COM : control mode status to HMI
	COM.HMI_OUTPUT_LOCAL_ACTIVE := INTERN.LOCAL_HMI;

	//--- EXC
	EXC.EXC_OUTPUT_FREQUENCY            := INTERN.FREQUENCY;
	EXC.EXC_OUTPUT_L1_N_VOLTAGE         := INTERN.L1_N_VOLTAGE;
	EXC.EXC_OUTPUT_L1_CURRENT           := INTERN.L1_CURRENT;
	EXC.EXC_OUTPUT_L1_ACTIVE_POWER      := INTERN.L1_ACTIVE_POWER;
	EXC.EXC_OUTPUT_L1_APPARENT_POWER    := INTERN.L1_APPARENT_POWER;
	EXC.EXC_OUTPUT_L1_REACTIVE_POWER    := INTERN.L1_REACTIVE_POWER;
	EXC.EXC_OUTPUT_L1_POWER_FACTOR      := INTERN.L1_POWER_FACTOR;
	EXC.EXC_OUTPUT_L1_VOLTAGE_THD       := INTERN.L1_VOLTAGE_THD;
	EXC.EXC_OUTPUT_L1_CURRENT_THD       := INTERN.L1_CURRENT_THD;
	EXC.EXC_OUTPUT_L1_MAX_LOAD          := INTERN.L1_MAX_LOAD;
	EXC.EXC_OUTPUT_INTERNAL_TEMPERATURE := INTERN.INTERNAL_TEMPERATURE;
	EXC.EXC_OUTPUT_ACTIVE_ENERGY        := INTERN.ACTIVE_ENERGY;
	// EXC.EXC_OUTPUT_DATA_VALID : not managed yet (no Modbus diagnostic)

	//--- COM : alarms to HMI
	COM.HMI_OUTPUT_ALARM_1_STATUS  := INTERN.ALARM_1;
	COM.HMI_OUTPUT_ALARM_2_STATUS  := INTERN.ALARM_2;
	COM.HMI_OUTPUT_ALARM_3_STATUS  := INTERN.ALARM_3;
	COM.HMI_OUTPUT_ALARM_4_STATUS  := INTERN.ALARM_4;
	COM.HMI_OUTPUT_ALARM_5_STATUS  := INTERN.ALARM_5;
	COM.HMI_OUTPUT_ALARM_6_STATUS  := INTERN.ALARM_6;
	COM.HMI_OUTPUT_ALARM_7_STATUS  := INTERN.ALARM_7;
	COM.HMI_OUTPUT_ALARM_8_STATUS  := INTERN.ALARM_8;
	COM.HMI_OUTPUT_ALARM_9_STATUS  := INTERN.ALARM_9;
	COM.HMI_OUTPUT_ALARM_10_STATUS := INTERN.ALARM_10;

	//--- COM : measures to HMI
	COM.HMI_OUTPUT_FREQUENCY.Real_value                 := INTERN.FREQUENCY;
	COM.HMI_OUTPUT_L1_L2_VOLTAGE.Real_value             := INTERN.L1_L2_VOLTAGE;
	COM.HMI_OUTPUT_L1_N_VOLTAGE.Real_value              := INTERN.L1_N_VOLTAGE;
	COM.HMI_OUTPUT_L1_CURRENT.Real_value                := INTERN.L1_CURRENT;
	COM.HMI_OUTPUT_L1_ACTIVE_POWER.Real_value           := INTERN.L1_ACTIVE_POWER;
	COM.HMI_OUTPUT_L1_APPARENT_POWER.Real_value         := INTERN.L1_APPARENT_POWER;
	COM.HMI_OUTPUT_L1_REACTIVE_POWER.Real_value         := INTERN.L1_REACTIVE_POWER;
	COM.HMI_OUTPUT_L1_CURRENT_PHASE_ANGLE.Real_value    := INTERN.L1_CURRENT_PHASE_ANGLE;
	COM.HMI_OUTPUT_L1_POWER_FACTOR.Real_value           := INTERN.L1_POWER_FACTOR;
	COM.HMI_OUTPUT_L1_VOLTAGE_THD.Real_value            := INTERN.L1_VOLTAGE_THD;
	COM.HMI_OUTPUT_L1_CURRENT_THD.Real_value            := INTERN.L1_CURRENT_THD;
	COM.HMI_OUTPUT_L1_MAX_LOAD.Real_value               := INTERN.L1_MAX_LOAD;
	COM.HMI_OUTPUT_L1_L2_VOLTAGE_PHASE_ANGLE.Real_value := INTERN.L1_L2_VOLTAGE_PHASE_ANGLE;
	COM.HMI_OUTPUT_L2_L3_VOLTAGE.Real_value             := INTERN.L2_L3_VOLTAGE;
	COM.HMI_OUTPUT_L2_N_VOLTAGE.Real_value              := INTERN.L2_N_VOLTAGE;
	COM.HMI_OUTPUT_L2_CURRENT.Real_value                := INTERN.L2_CURRENT;
	COM.HMI_OUTPUT_L2_ACTIVE_POWER.Real_value           := INTERN.L2_ACTIVE_POWER;
	COM.HMI_OUTPUT_L2_APPARENT_POWER.Real_value         := INTERN.L2_APPARENT_POWER;
	COM.HMI_OUTPUT_L2_REACTIVE_POWER.Real_value         := INTERN.L2_REACTIVE_POWER;
	COM.HMI_OUTPUT_L2_CURRENT_PHASE_ANGLE.Real_value    := INTERN.L2_CURRENT_PHASE_ANGLE;
	COM.HMI_OUTPUT_L2_POWER_FACTOR.Real_value           := INTERN.L2_POWER_FACTOR;
	COM.HMI_OUTPUT_L2_VOLTAGE_THD.Real_value            := INTERN.L2_VOLTAGE_THD;
	COM.HMI_OUTPUT_L2_CURRENT_THD.Real_value            := INTERN.L2_CURRENT_THD;
	COM.HMI_OUTPUT_L2_MAX_LOAD.Real_value               := INTERN.L2_MAX_LOAD;
	COM.HMI_OUTPUT_L1_L3_VOLTAGE_PHASE_ANGLE.Real_value := INTERN.L1_L3_VOLTAGE_PHASE_ANGLE;
	COM.HMI_OUTPUT_L3_L1_VOLTAGE.Real_value             := INTERN.L3_L1_VOLTAGE;
	COM.HMI_OUTPUT_L3_N_VOLTAGE.Real_value              := INTERN.L3_N_VOLTAGE;
	COM.HMI_OUTPUT_L3_CURRENT.Real_value                := INTERN.L3_CURRENT;
	COM.HMI_OUTPUT_L3_ACTIVE_POWER.Real_value           := INTERN.L3_ACTIVE_POWER;
	COM.HMI_OUTPUT_L3_APPARENT_POWER.Real_value         := INTERN.L3_APPARENT_POWER;
	COM.HMI_OUTPUT_L3_REACTIVE_POWER.Real_value         := INTERN.L3_REACTIVE_POWER;
	COM.HMI_OUTPUT_L3_CURRENT_PHASE_ANGLE.Real_value    := INTERN.L3_CURRENT_PHASE_ANGLE;
	COM.HMI_OUTPUT_L3_POWER_FACTOR.Real_value           := INTERN.L3_POWER_FACTOR;
	COM.HMI_OUTPUT_L3_VOLTAGE_THD.Real_value            := INTERN.L3_VOLTAGE_THD;
	COM.HMI_OUTPUT_L3_CURRENT_THD.Real_value            := INTERN.L3_CURRENT_THD;
	COM.HMI_OUTPUT_L3_MAX_LOAD.Real_value               := INTERN.L3_MAX_LOAD;
	COM.HMI_OUTPUT_INTERNAL_TEMPERATURE.Real_value      := INTERN.INTERNAL_TEMPERATURE;
	COM.HMI_OUTPUT_ACTIVE_ENERGY.Real_value             := INTERN.ACTIVE_ENERGY;
	COM.HMI_OUTPUT_APPARENT_ENERGY.Real_value           := INTERN.APPARENT_ENERGY;
	COM.HMI_OUTPUT_REACTIVE_ENERGY.Real_value           := INTERN.REACTIVE_ENERGY;
	COM.HMI_OUTPUT_TOTAL_ACTIVE_POWER.Real_value        := INTERN.TOTAL_ACTIVE_POWER;
	COM.HMI_OUTPUT_TOTAL_APPARENT_POWER.Real_value      := INTERN.TOTAL_APPARENT_POWER;
	COM.HMI_OUTPUT_TOTAL_REACTIVE_POWER.Real_value      := INTERN.TOTAL_REACTIVE_POWER;
	COM.HMI_OUTPUT_ALL_PHASE_POWER_FACTOR.Real_value    := INTERN.ALL_PHASE_POWER_FACTOR;


                
END_FUNCTION_BLOCK

FUNCTION_BLOCK FB_INST_DIP1500
  VAR_IN_OUT
    PA : DUT_PA_DIP1500;  (* Parameters (persistent, GVL_PA) *)
    COM : DUT_COM_DIP1500;  (* Communication : Modbus RTU (COM_), HMI PanelView (HMI_) *)
    EXC : DUT_EXC_DIP1500;  (* Exchanges : other equipment (EXC_), functional units (UPI_) *)
    IO : DUT_IO_DIP1500;  (* Wired PLC I/O *)
  END_VAR
  VAR
    INTERN : DUT_INT_DIP1500;  (* Internal variables *)
    TON_PULSE : TON;  (* Square wave timer *)
    TOF_CMD_WINDOW : TOF;  (* Command write window *)
    R_TRIG_FLASH : R_TRIG;  (* Flash save request edge *)
    TP_FLASH : TP;  (* Flash save pulse *)
  END_VAR

                  
//==============================================================================
// FB_INST_DIP1500
// Kamoer DIP1500 peristaltic pump, Modbus RTU, 32-bit low word first (CDAB)
// 1. INPUTS     : requests, control mode, command source, equipment feedback -> INTERN
// 2. PROCESSING : on INTERN only
// 3. OUTPUTS    : INTERN -> COM / IO / EXC
// Parameters    : pump configuration in PA (persistent), changed from the HMI in local HMI
// Control mode  : local HMI (individual or global) > auto (functional units)
//==============================================================================

//------------------------------------------------------------------------------
// 1. INPUTS
//------------------------------------------------------------------------------
	//--- Control mode requests (HMI, global HMI local from UPI_LOCAL_HMI)
	INTERN.HMI_LOCAL_REQUEST := COM.HMI_INPUT_LOCAL_REQUEST;
	INTERN.HMI_AUTO_REQUEST  := COM.HMI_INPUT_AUTO_REQUEST;
	INTERN.GLOBAL_LOCAL_HMI  := EXC.UPI_INPUT_GLOBAL_LOCAL_HMI;

	//--- Control mode
	// Individual memory : set by the local request, reset by the auto request (auto wins if both)
	IF INTERN.HMI_LOCAL_REQUEST THEN
		INTERN.LOCAL_HMI_INDIVIDUAL := TRUE;
	END_IF
	IF INTERN.HMI_AUTO_REQUEST THEN
		INTERN.LOCAL_HMI_INDIVIDUAL := FALSE;
	END_IF

	// Resulting mode : HMI local (individual OR global), otherwise auto
	INTERN.LOCAL_HMI := INTERN.LOCAL_HMI_INDIVIDUAL OR INTERN.GLOBAL_LOCAL_HMI;
	INTERN.AUTO      := NOT INTERN.LOCAL_HMI;
	
	//--- Command source : local HMI > auto (UPI)
	IF INTERN.LOCAL_HMI THEN
		INTERN.CMD_RUN            := COM.HMI_INPUT_MOTOR_START_STOP;
		INTERN.CMD_CLOCKWISE      := COM.HMI_INPUT_MOTOR_DIRECTION;
		INTERN.CMD_VOLUME_MODE    := COM.HMI_INPUT_OPERATION_MODE;
		INTERN.CMD_SPEED          := COM.HMI_INPUT_MOTOR_SPEED.Real_value;
		INTERN.CMD_RUN_SETPOINT   := COM.HMI_INPUT_RUN_TIME_OR_VOLUME_SETPOINT.Real_value;
		INTERN.PARAM_WRITE_ENABLE := COM.HMI_INPUT_PARAM_WRITE_ENABLE;
		INTERN.FLASH_SAVE_REQUEST := COM.HMI_INPUT_FLASH_SAVE;
	ELSE
		// Auto : functional units (UPI)
		INTERN.CMD_RUN            := EXC.UPI_INPUT_RUN;
		INTERN.CMD_CLOCKWISE      := EXC.UPI_INPUT_CLOCKWISE;
		INTERN.CMD_VOLUME_MODE    := EXC.UPI_INPUT_VOLUME_MODE;
		INTERN.CMD_SPEED          := EXC.UPI_INPUT_SPEED;
		INTERN.CMD_RUN_SETPOINT   := EXC.UPI_INPUT_RUN_SETPOINT;
		INTERN.PARAM_WRITE_ENABLE := FALSE;                        // configuration is never written in auto
		INTERN.FLASH_SAVE_REQUEST := FALSE;
	END_IF
	
	//--- Parameter source : values typed on the HMI in local HMI (nothing in auto)
	IF INTERN.LOCAL_HMI THEN
		INTERN.SRC_MAX_MOTOR_SPEED         := COM.HMI_INPUT_MAX_MOTOR_SPEED.Real_value;
		INTERN.SRC_CALIBRATION_COEFFICIENT := COM.HMI_INPUT_FLOW_RATE_OR_SPEED_CALIBRATION_COEFFICIENT.Real_value;
		INTERN.SRC_FOOT_SWITCH_INPUT_MODE  := COM.HMI_INPUT_FOOT_SWITCH_INPUT_MODE;
		INTERN.SRC_LIQUID_LEVEL_INPUT_MODE := COM.HMI_INPUT_LIQUID_LEVEL_INPUT_MODE;
		INTERN.SRC_STATE_OUTPUT_MODE       := COM.HMI_INPUT_STATE_OUTPUT_MODE;
		INTERN.SRC_COMMUNICATION_ADDRESS   := COM.HMI_INPUT_COMMUNICATION_ADDRESS;
		INTERN.SRC_BAUD_RATE_INDEX         := COM.HMI_INPUT_BAUD_RATE_INDEX;
	END_IF
	
	//--- COM : input registers 0x3001..0x3005
	INTERN.FBK_FIRMWARE_VERSION := COM.COM_INPUT_IR[0];
	INTERN.FBK_HARDWARE_VERSION := COM.COM_INPUT_IR[1];
	INTERN.FBK_TEMPERATURE      := COM.COM_INPUT_IR[2];
	INTERN.FBK_LEVEL_ALARM      := COM.COM_INPUT_IR[3];
	INTERN.FBK_DIGITAL_OUTPUT   := COM.COM_INPUT_IR[4];
	
	//--- COM : run counters 0x4007..0x400A (format depends on mode)
	IF INTERN.CMD_VOLUME_MODE THEN
		// Volume mode : 32-bit REAL (ml)
		INTERN.FBK_RUN_ACTUAL := FNC_WORDS_TO_REAL(High_word := COM.COM_INPUT_HR_COUNTERS[1], Low_word := COM.COM_INPUT_HR_COUNTERS[0]);
		INTERN.FBK_RUN_TOTAL  := FNC_WORDS_TO_REAL(High_word := COM.COM_INPUT_HR_COUNTERS[3], Low_word := COM.COM_INPUT_HR_COUNTERS[2]);
	ELSE
		// Time mode : 32-bit UDINT (ms)
		INTERN.UDINT_TEMP     := SHL(WORD_TO_UDINT(COM.COM_INPUT_HR_COUNTERS[1]), 16) OR WORD_TO_UDINT(COM.COM_INPUT_HR_COUNTERS[0]);
		INTERN.FBK_RUN_ACTUAL := UDINT_TO_REAL(INTERN.UDINT_TEMP);
		INTERN.UDINT_TEMP     := SHL(WORD_TO_UDINT(COM.COM_INPUT_HR_COUNTERS[3]), 16) OR WORD_TO_UDINT(COM.COM_INPUT_HR_COUNTERS[2]);
		INTERN.FBK_RUN_TOTAL  := UDINT_TO_REAL(INTERN.UDINT_TEMP);
	END_IF
	
	
//------------------------------------------------------------------------------
// 2. PROCESSING
//------------------------------------------------------------------------------
	//--- Parameters (PA) : a value changed on the HMI (local HMI) is saved in PA
	// PA is persistent : it keeps its value after a restart or a download. Default = declaration value.
	// The cycle where the mode changes is ignored, so switching mode never overwrites PA.
	INTERN.SOURCE_CHANGED := INTERN.LOCAL_HMI <> INTERN.PREV_LOCAL_HMI;
	INTERN.PREV_LOCAL_HMI := INTERN.LOCAL_HMI;
	
	IF NOT INTERN.SOURCE_CHANGED THEN
		IF INTERN.SRC_MAX_MOTOR_SPEED <> INTERN.PREV_SRC_MAX_MOTOR_SPEED THEN
			PA.MAX_MOTOR_SPEED := INTERN.SRC_MAX_MOTOR_SPEED;
		END_IF
		IF INTERN.SRC_CALIBRATION_COEFFICIENT <> INTERN.PREV_SRC_CALIBRATION_COEFFICIENT THEN
			PA.CALIBRATION_COEFFICIENT := INTERN.SRC_CALIBRATION_COEFFICIENT;
		END_IF
		IF INTERN.SRC_FOOT_SWITCH_INPUT_MODE <> INTERN.PREV_SRC_FOOT_SWITCH_INPUT_MODE THEN
			PA.FOOT_SWITCH_INPUT_MODE := INTERN.SRC_FOOT_SWITCH_INPUT_MODE;
		END_IF
		IF INTERN.SRC_LIQUID_LEVEL_INPUT_MODE <> INTERN.PREV_SRC_LIQUID_LEVEL_INPUT_MODE THEN
			PA.LIQUID_LEVEL_INPUT_MODE := INTERN.SRC_LIQUID_LEVEL_INPUT_MODE;
		END_IF
		IF INTERN.SRC_STATE_OUTPUT_MODE <> INTERN.PREV_SRC_STATE_OUTPUT_MODE THEN
			PA.STATE_OUTPUT_MODE := INTERN.SRC_STATE_OUTPUT_MODE;
		END_IF
		IF INTERN.SRC_COMMUNICATION_ADDRESS <> INTERN.PREV_SRC_COMMUNICATION_ADDRESS THEN
			PA.COMMUNICATION_ADDRESS := INTERN.SRC_COMMUNICATION_ADDRESS;
		END_IF
		IF INTERN.SRC_BAUD_RATE_INDEX <> INTERN.PREV_SRC_BAUD_RATE_INDEX THEN
			PA.BAUD_RATE_INDEX := INTERN.SRC_BAUD_RATE_INDEX;
		END_IF
	END_IF
	
	INTERN.PREV_SRC_MAX_MOTOR_SPEED         := INTERN.SRC_MAX_MOTOR_SPEED;
	INTERN.PREV_SRC_CALIBRATION_COEFFICIENT := INTERN.SRC_CALIBRATION_COEFFICIENT;
	INTERN.PREV_SRC_FOOT_SWITCH_INPUT_MODE  := INTERN.SRC_FOOT_SWITCH_INPUT_MODE;
	INTERN.PREV_SRC_LIQUID_LEVEL_INPUT_MODE := INTERN.SRC_LIQUID_LEVEL_INPUT_MODE;
	INTERN.PREV_SRC_STATE_OUTPUT_MODE       := INTERN.SRC_STATE_OUTPUT_MODE;
	INTERN.PREV_SRC_COMMUNICATION_ADDRESS   := INTERN.SRC_COMMUNICATION_ADDRESS;
	INTERN.PREV_SRC_BAUD_RATE_INDEX         := INTERN.SRC_BAUD_RATE_INDEX;
	
	//--- Parameters used by the pump : always from PA
	INTERN.CMD_MAX_SPEED      := PA.MAX_MOTOR_SPEED;
	INTERN.CMD_CALIB_COEF     := PA.CALIBRATION_COEFFICIENT;
	INTERN.CMD_FOOT_MODE      := PA.FOOT_SWITCH_INPUT_MODE;
	INTERN.CMD_LEVEL_MODE     := PA.LIQUID_LEVEL_INPUT_MODE;
	INTERN.CMD_STATE_OUT_MODE := PA.STATE_OUTPUT_MODE;
	INTERN.CMD_ADDRESS        := PA.COMMUNICATION_ADDRESS;
	INTERN.CMD_BAUD_INDEX     := PA.BAUD_RATE_INDEX;
	
	//--- Parameter validity
	INTERN.PARAM_VALID := (WORD_TO_UINT(INTERN.CMD_ADDRESS) >= 1) AND (WORD_TO_UINT(INTERN.CMD_ADDRESS) <= 31)
	                      AND (WORD_TO_UINT(INTERN.CMD_BAUD_INDEX) <= 7)
	                      AND (INTERN.CMD_MAX_SPEED > 0.0) AND (INTERN.CMD_CALIB_COEF > 0.0);

	//--- Flash save : 1 s pulse on rising edge, only with valid parameters
	R_TRIG_FLASH(CLK := INTERN.FLASH_SAVE_REQUEST);
	TP_FLASH(IN := R_TRIG_FLASH.Q AND INTERN.PARAM_VALID, PT := T#1S);
	INTERN.CMD_SAVE_FLASH := TP_FLASH.Q;
	
	//--- Write triggers (rising edge channels)
	// Square wave 500 ms : each rising edge = one write request
	TON_PULSE(IN := NOT TON_PULSE.Q, PT := T#250MS);
	IF TON_PULSE.Q THEN
		INTERN.PULSE_500MS := NOT INTERN.PULSE_500MS;
	END_IF
	
	// Command trigger : automatic, 3 s of edges after any command change
	INTERN.CMD_CHANGED := (INTERN.CMD_RUN <> INTERN.PREV_RUN) OR (INTERN.CMD_CLOCKWISE <> INTERN.PREV_CLOCKWISE)
	                      OR (INTERN.CMD_VOLUME_MODE <> INTERN.PREV_VOLUME_MODE) OR (INTERN.CMD_SAVE_FLASH <> INTERN.PREV_SAVE_FLASH)
	                      OR (INTERN.CMD_SPEED <> INTERN.PREV_SPEED) OR (INTERN.CMD_MAX_SPEED <> INTERN.PREV_MAX_SPEED)
	                      OR (INTERN.CMD_RUN_SETPOINT <> INTERN.PREV_RUN_SETPOINT);
	INTERN.PREV_RUN          := INTERN.CMD_RUN;
	INTERN.PREV_CLOCKWISE    := INTERN.CMD_CLOCKWISE;
	INTERN.PREV_VOLUME_MODE  := INTERN.CMD_VOLUME_MODE;
	INTERN.PREV_SAVE_FLASH   := INTERN.CMD_SAVE_FLASH;
	INTERN.PREV_SPEED        := INTERN.CMD_SPEED;
	INTERN.PREV_MAX_SPEED    := INTERN.CMD_MAX_SPEED;
	INTERN.PREV_RUN_SETPOINT := INTERN.CMD_RUN_SETPOINT;
	
	TOF_CMD_WINDOW(IN := INTERN.CMD_CHANGED, PT := T#3S);
	INTERN.CMD_WINDOW  := TOF_CMD_WINDOW.Q;
	INTERN.CMD_TRIGGER := INTERN.CMD_WINDOW AND (INTERN.CMD_MAX_SPEED > 0.0) AND INTERN.PULSE_500MS;
	
	// Configuration trigger : only while writing is enabled and parameters are valid
	INTERN.CONFIG_TRIGGER := INTERN.PARAM_WRITE_ENABLE AND INTERN.PARAM_VALID AND INTERN.PULSE_500MS;
	
	
//------------------------------------------------------------------------------
// 3. OUTPUTS
//------------------------------------------------------------------------------
	//--- COM : control mode status to HMI
	COM.HMI_OUTPUT_LOCAL_ACTIVE := INTERN.LOCAL_HMI;
	
	//--- COM : Modbus RTU coils
	COM.COM_OUTPUT_COILS[0] := INTERN.CMD_RUN;           // 0x0001
	COM.COM_OUTPUT_COILS[1] := INTERN.CMD_CLOCKWISE;     // 0x0002
	COM.COM_OUTPUT_COILS[2] := INTERN.CMD_SAVE_FLASH;    // 0x0003
	COM.COM_OUTPUT_COILS[3] := INTERN.CMD_VOLUME_MODE;   // 0x0004
	
	//--- COM : Modbus RTU holding registers and write triggers
	// Command registers 0x4001..0x4006 (sent on the command trigger)
	FNC_REAL_TO_WORDS(Real_value := INTERN.CMD_SPEED,     High_word => COM.COM_OUTPUT_HR_CMD[1], Low_word => COM.COM_OUTPUT_HR_CMD[0]);   // 0x4001-4002
	FNC_REAL_TO_WORDS(Real_value := INTERN.CMD_MAX_SPEED, High_word => COM.COM_OUTPUT_HR_CMD[3], Low_word => COM.COM_OUTPUT_HR_CMD[2]);   // 0x4003-4004
	IF INTERN.CMD_VOLUME_MODE THEN
		// Run setpoint 0x4005-4006, volume mode : 32-bit REAL (ml)
		FNC_REAL_TO_WORDS(Real_value := INTERN.CMD_RUN_SETPOINT, High_word => COM.COM_OUTPUT_HR_CMD[5], Low_word => COM.COM_OUTPUT_HR_CMD[4]);
	ELSE
		// Run setpoint 0x4005-4006, time mode : 32-bit UDINT (ms)
		INTERN.UDINT_TEMP        := REAL_TO_UDINT(MAX(INTERN.CMD_RUN_SETPOINT, 0.0));
		COM.COM_OUTPUT_HR_CMD[4] := UDINT_TO_WORD(INTERN.UDINT_TEMP);
		COM.COM_OUTPUT_HR_CMD[5] := UDINT_TO_WORD(SHR(INTERN.UDINT_TEMP, 16));
	END_IF
	
	// Configuration registers 0x400B..0x4011 (sent on the configuration trigger), updated only while enabled and valid
	IF INTERN.PARAM_WRITE_ENABLE AND INTERN.PARAM_VALID THEN
		FNC_REAL_TO_WORDS(Real_value := INTERN.CMD_CALIB_COEF, High_word => COM.COM_OUTPUT_HR_CONFIG[1], Low_word => COM.COM_OUTPUT_HR_CONFIG[0]);   // 0x400B-400C
		COM.COM_OUTPUT_HR_CONFIG[2] := INTERN.CMD_FOOT_MODE;        // 0x400D
		COM.COM_OUTPUT_HR_CONFIG[3] := INTERN.CMD_LEVEL_MODE;       // 0x400E
		COM.COM_OUTPUT_HR_CONFIG[4] := INTERN.CMD_STATE_OUT_MODE;   // 0x400F
		COM.COM_OUTPUT_HR_CONFIG[5] := INTERN.CMD_ADDRESS;          // 0x4010
		COM.COM_OUTPUT_HR_CONFIG[6] := INTERN.CMD_BAUD_INDEX;       // 0x4011
	END_IF
	
	// Write triggers
	COM.COM_OUTPUT_CMD_TRIGGER    := INTERN.CMD_TRIGGER;
	COM.COM_OUTPUT_CONFIG_TRIGGER := INTERN.CONFIG_TRIGGER;
	
	//--- COM : feedback to HMI
	COM.HMI_OUTPUT_FIRMWARE_VERSION                          := INTERN.FBK_FIRMWARE_VERSION;
	COM.HMI_OUTPUT_HARDWARE_VERSION                          := INTERN.FBK_HARDWARE_VERSION;
	COM.HMI_OUTPUT_TEMPERATURE                               := INTERN.FBK_TEMPERATURE;
	COM.HMI_OUTPUT_FLOAT_LEVEL_ALARM                         := INTERN.FBK_LEVEL_ALARM;
	COM.HMI_OUTPUT_DIGITAL_OUTPUT_VALUE                      := INTERN.FBK_DIGITAL_OUTPUT;
	COM.HMI_OUTPUT_REAL_TIME_RUN_TIME_OR_VOLUME.Real_value   := INTERN.FBK_RUN_ACTUAL;
	COM.HMI_OUTPUT_ACCUMULATED_RUN_TIME_OR_VOLUME.Real_value := INTERN.FBK_RUN_TOTAL;


                
END_FUNCTION_BLOCK

FUNCTION_BLOCK FB_INST_DOSENSOR
  VAR_IN_OUT
    PA : DUT_PA_DOSENSOR;  (* Parameters (persistent, GVL_PA) *)
    COM : DUT_COM_DOSENSOR;  (* Communication : Modbus RTU (COM_), HMI PanelView (HMI_) *)
    EXC : DUT_EXC_DOSENSOR;  (* Exchanges : other equipment (EXC_), functional units (UPI_) *)
    IO : DUT_IO_DOSENSOR;  (* Wired PLC I/O *)
  END_VAR
  VAR
    INTERN : DUT_INT_DOSENSOR;  (* Internal variables *)
    TP_CALIB_HIGH : TP;  (* High calibration pulse *)
    TP_CALIB_LOW : TP;  (* Low calibration pulse *)
    TP_CALIB_DONE : TP;  (* Calibration done message *)
  END_VAR

                  
//==============================================================================
// FB_INST_DOSENSOR
// Dissolved oxygen sensor, analog signal + fault input + 2 calibration outputs
// 1. INPUTS     : requests, control mode, command source, equipment feedback -> INTERN
// 2. PROCESSING : on INTERN only
// 3. OUTPUTS    : INTERN -> COM / IO / EXC
// Control mode  : local HMI (individual or global) > auto (functional units)
//==============================================================================

//------------------------------------------------------------------------------
// 1. INPUTS
//------------------------------------------------------------------------------
	//--- Control mode requests (HMI, global HMI local from UPI_LOCAL_HMI)
	INTERN.HMI_LOCAL_REQUEST := COM.HMI_INPUT_LOCAL_REQUEST;
	INTERN.HMI_AUTO_REQUEST  := COM.HMI_INPUT_AUTO_REQUEST;
	INTERN.GLOBAL_LOCAL_HMI  := EXC.UPI_INPUT_GLOBAL_LOCAL_HMI;

	//--- Control mode
	// Individual memory : set by the local request, reset by the auto request (auto wins if both)
	IF INTERN.HMI_LOCAL_REQUEST THEN
		INTERN.LOCAL_HMI_INDIVIDUAL := TRUE;
	END_IF
	IF INTERN.HMI_AUTO_REQUEST THEN
		INTERN.LOCAL_HMI_INDIVIDUAL := FALSE;
	END_IF

	// Resulting mode : HMI local (individual OR global), otherwise auto
	INTERN.LOCAL_HMI := INTERN.LOCAL_HMI_INDIVIDUAL OR INTERN.GLOBAL_LOCAL_HMI;
	INTERN.AUTO      := NOT INTERN.LOCAL_HMI;

	//--- Command source : calibration requests (local HMI > auto)
	IF INTERN.LOCAL_HMI THEN
		INTERN.CALIB_HIGH_REQUEST := COM.HMI_INPUT_CALIBRATION_HIGH;
		INTERN.CALIB_LOW_REQUEST  := COM.HMI_INPUT_CALIBRATION_LOW;
	ELSE
		// Auto : functional units (UPI)
		INTERN.CALIB_HIGH_REQUEST := FALSE;
		INTERN.CALIB_LOW_REQUEST  := FALSE;
	END_IF

	//--- IO
	INTERN.SIGNAL_RAW := IO.INPUT_SIGNAL;
	INTERN.FAULT      := IO.INPUT_SENSOR_FAULT;


//------------------------------------------------------------------------------
// 2. PROCESSING
//------------------------------------------------------------------------------
	//--- Signal scaling
	INTERN.SIGNAL := (DWORD_TO_REAL(INTERN.SIGNAL_RAW * 40) / 65535) - 8;

	//--- Calibration : 1 s pulse to the sensor, 5 s "done" message
	TP_CALIB_HIGH(IN := INTERN.CALIB_HIGH_REQUEST, PT := T#1S);
	TP_CALIB_LOW(IN := INTERN.CALIB_LOW_REQUEST, PT := T#1S);
	TP_CALIB_DONE(IN := TP_CALIB_HIGH.Q OR TP_CALIB_LOW.Q, PT := T#5S);

	INTERN.CALIB_HIGH := TP_CALIB_HIGH.Q;
	INTERN.CALIB_LOW  := TP_CALIB_LOW.Q;
	INTERN.CALIB_DONE := TP_CALIB_DONE.Q;


//------------------------------------------------------------------------------
// 3. OUTPUTS
//------------------------------------------------------------------------------
	//--- COM : control mode status to HMI
	COM.HMI_OUTPUT_LOCAL_ACTIVE := INTERN.LOCAL_HMI;

	//--- EXC
	EXC.EXC_OUTPUT_SIGNAL := INTERN.SIGNAL;

	//--- IO
	IO.OUTPUT_CALIBRATION_HIGH := INTERN.CALIB_HIGH;
	IO.OUTPUT_CALIBRATION_LOW  := INTERN.CALIB_LOW;

	//--- COM : feedback to HMI
	COM.HMI_OUTPUT_SIGNAL.Real_value := INTERN.SIGNAL;
	COM.HMI_OUTPUT_FAULT             := INTERN.FAULT;
	COM.HMI_OUTPUT_CALIBRATION_DONE  := INTERN.CALIB_DONE;


                
END_FUNCTION_BLOCK

FUNCTION_BLOCK FB_UPI_LOCAL_HMI
  VAR_IN_OUT
    COM : DUT_COM_UPI_LOCAL_HMI;  (* Requests and status with the HMI *)
    EXC : DUT_EXC_UPI_LOCAL_HMI;  (* Status to equipment *)
  END_VAR
  VAR
    INTERN : DUT_INT_UPI_LOCAL_HMI;  (* Internal variables *)
  END_VAR

                  
//==============================================================================
// FB_UPI_LOCAL_HMI
// Global HMI local mode for every equipment
// Set by the HMI local request, reset by the HMI auto request (pulse or maintained, auto wins)
// The equipment read this status through GFC_EXC and report their own local status themselves
//==============================================================================

//------------------------------------------------------------------------------
// 1. INPUTS
//------------------------------------------------------------------------------
	INTERN.LOCAL_REQUEST := COM.HMI_INPUT_LOCAL_REQUEST;
	INTERN.AUTO_REQUEST  := COM.HMI_INPUT_AUTO_REQUEST;


//------------------------------------------------------------------------------
// 2. PROCESSING
//------------------------------------------------------------------------------
	IF INTERN.LOCAL_REQUEST THEN
		INTERN.LOCAL_ACTIVE := TRUE;
	END_IF
	IF INTERN.AUTO_REQUEST THEN
		INTERN.LOCAL_ACTIVE := FALSE;
	END_IF


//------------------------------------------------------------------------------
// 3. OUTPUTS
//------------------------------------------------------------------------------
	//--- EXC : to every equipment (through GFC_EXC)
	EXC.UPI_OUTPUT_LOCAL_ACTIVE := INTERN.LOCAL_ACTIVE;

	//--- COM : status
	COM.HMI_OUTPUT_LOCAL_ACTIVE := INTERN.LOCAL_ACTIVE;


                
END_FUNCTION_BLOCK

FUNCTION FC_EXC_UPI_LOCAL_HMI_ADM100W : BOOL
  VAR_IN_OUT
    EXC_UPI_LOCAL_HMI : DUT_EXC_UPI_LOCAL_HMI;  (* Exchanges of the UPI_LOCAL_HMI instance *)
    EXC_ADM100W : DUT_EXC_ADM100W;  (* Exchanges of the ADM100W instance *)
  END_VAR

                  
//==============================================================================
// FC_EXC_UPI_LOCAL_HMI_ADM100W
// Exchanges between one UPI_LOCAL_HMI instance and one ADM100W instance
// Called in GFC_EXC, once per pair of instances, with their GVL_EXC variables
// Simple copies only, no conversion
//==============================================================================

//--- UPI_LOCAL_HMI -> ADM100W
EXC_ADM100W.UPI_INPUT_GLOBAL_LOCAL_HMI := EXC_UPI_LOCAL_HMI.UPI_OUTPUT_LOCAL_ACTIVE;

FC_EXC_UPI_LOCAL_HMI_ADM100W := TRUE;

                
END_FUNCTION

FUNCTION FC_EXC_UPI_LOCAL_HMI_DIP1500 : BOOL
  VAR_IN_OUT
    EXC_UPI_LOCAL_HMI : DUT_EXC_UPI_LOCAL_HMI;  (* Exchanges of the UPI_LOCAL_HMI instance *)
    EXC_DIP1500 : DUT_EXC_DIP1500;  (* Exchanges of the DIP1500 instance *)
  END_VAR

                  
//==============================================================================
// FC_EXC_UPI_LOCAL_HMI_DIP1500
// Exchanges between one UPI_LOCAL_HMI instance and one DIP1500 instance
// Called in GFC_EXC, once per pair of instances, with their GVL_EXC variables
// Simple copies only, no conversion
//==============================================================================

//--- UPI_LOCAL_HMI -> DIP1500
EXC_DIP1500.UPI_INPUT_GLOBAL_LOCAL_HMI := EXC_UPI_LOCAL_HMI.UPI_OUTPUT_LOCAL_ACTIVE;

FC_EXC_UPI_LOCAL_HMI_DIP1500 := TRUE;

                
END_FUNCTION

FUNCTION FC_EXC_UPI_LOCAL_HMI_DOSENSOR : BOOL
  VAR_IN_OUT
    EXC_UPI_LOCAL_HMI : DUT_EXC_UPI_LOCAL_HMI;  (* Exchanges of the UPI_LOCAL_HMI instance *)
    EXC_DOSENSOR : DUT_EXC_DOSENSOR;  (* Exchanges of the DOSENSOR instance *)
  END_VAR

                  
//==============================================================================
// FC_EXC_UPI_LOCAL_HMI_DOSENSOR
// Exchanges between one UPI_LOCAL_HMI instance and one DOSENSOR instance
// Called in GFC_EXC, once per pair of instances, with their GVL_EXC variables
// Simple copies only, no conversion
//==============================================================================

//--- UPI_LOCAL_HMI -> DOSENSOR
EXC_DOSENSOR.UPI_INPUT_GLOBAL_LOCAL_HMI := EXC_UPI_LOCAL_HMI.UPI_OUTPUT_LOCAL_ACTIVE;

FC_EXC_UPI_LOCAL_HMI_DOSENSOR := TRUE;

                
END_FUNCTION

FUNCTION FNC_REAL_TO_WORDS : BOOL
  VAR_INPUT
    Real_value : REAL;  (* Value to split *)
  END_VAR
  VAR_OUTPUT
    High_word : WORD;  (* Most significant word *)
    Low_word : WORD;  (* Least significant word *)
  END_VAR
  VAR
    Conversion : DUT_Union_Real_Word;  (* REAL / 2 WORD overlay *)
  END_VAR

                  
//==============================================================================
// FNC_REAL_TO_WORDS
// REAL (IEEE 754) -> two Modbus words
// Call: FNC_REAL_TO_WORDS(Real_value := x, High_word => ..., Low_word => ...);
//==============================================================================

Conversion.Real_value := Real_value;
Low_word  := Conversion.Word_value[0];
High_word := Conversion.Word_value[1];
FNC_REAL_TO_WORDS := TRUE;

                
END_FUNCTION

FUNCTION FNC_WORDS_TO_REAL : REAL
  VAR_INPUT
    High_word : WORD;  (* Most significant word *)
    Low_word : WORD;  (* Least significant word *)
  END_VAR
  VAR
    Conversion : DUT_Union_Real_Word;  (* REAL / 2 WORD overlay *)
  END_VAR

                  
//==============================================================================
// FNC_WORDS_TO_REAL
// Two Modbus words -> REAL (IEEE 754)
// ABCD device: High_word = lower address, CDAB device: Low_word = lower address
//==============================================================================

Conversion.Word_value[0] := Low_word;
Conversion.Word_value[1] := High_word;
FNC_WORDS_TO_REAL := Conversion.Real_value;

                
END_FUNCTION

FUNCTION_BLOCK GFB_INST
  VAR
    FB_ADM100W_1 : FB_INST_ADM100W;  (* Trumeter ADM100W power meter *)
    FB_DOSENSOR_1 : FB_INST_DOSENSOR;  (* Dissolved oxygen sensor *)
    FB_DIP1500_1 : FB_INST_DIP1500;  (* Kamoer DIP1500 peristaltic pump *)
  END_VAR

                  
//==============================================================================
// GFB_INST
// Calls every equipment instance
// One block per equipment, all interfaces connected
//==============================================================================

//--- ADM100W_1 : Trumeter ADM100W power meter
FB_ADM100W_1(
	PA  := GVL_PA.PA_ADM100W_1,
	COM := GVL_COM.COM_ADM100W_1,
	EXC := GVL_EXC.EXC_ADM100W_1,
	IO  := GVL_IO.IO_ADM100W_1);

//--- DOSENSOR_1 : Dissolved oxygen sensor
FB_DOSENSOR_1(
	PA  := GVL_PA.PA_DOSENSOR_1,
	COM := GVL_COM.COM_DOSENSOR_1,
	EXC := GVL_EXC.EXC_DOSENSOR_1,
	IO  := GVL_IO.IO_DOSENSOR_1);

//--- DIP1500_1 : Kamoer DIP1500 peristaltic pump
FB_DIP1500_1(
	PA  := GVL_PA.PA_DIP1500_1,
	COM := GVL_COM.COM_DIP1500_1,
	EXC := GVL_EXC.EXC_DIP1500_1,
	IO  := GVL_IO.IO_DIP1500_1);

                
END_FUNCTION_BLOCK

FUNCTION_BLOCK GFB_UPI
  VAR
    FB_UPI_LOCAL_HMI_1 : FB_UPI_LOCAL_HMI;  (* Global HMI local mode *)
  END_VAR

                  
//==============================================================================
// GFB_UPI
// Calls every functional unit (UPI)
// Runs before GFB_INST, results go to the equipment through GFC_EXC
//==============================================================================

//--- UPI_LOCAL_HMI : Global HMI local mode
FB_UPI_LOCAL_HMI_1(
	COM := GVL_COM.COM_UPI_LOCAL_HMI,
	EXC := GVL_EXC.EXC_UPI_LOCAL_HMI);


                
END_FUNCTION_BLOCK

FUNCTION GFC_COM_IN : BOOL

                  
//==============================================================================
// GFC_COM_IN
// Modbus (GVL_MODBUS) -> GVL_COM : RTU equipment, HMI
// Simple copies only, no conversion (conversions are done in the FBs)
//==============================================================================

//------------------------------------------------------------------------------
// COM : Modbus RTU, from equipment
//------------------------------------------------------------------------------
	//--- ADM100W_1
	GVL_COM.COM_ADM100W_1.COM_INPUT_IR    := GVL_MODBUS.ADM100W_InputRegisters;   // Input registers 0..87
	GVL_COM.COM_ADM100W_1.COM_INPUT_COILS := GVL_MODBUS.ADM100W_Alarms;           // Coils 0..9 (alarms)

	//--- DIP1500_1
	GVL_COM.COM_DIP1500_1.COM_INPUT_IR          := GVL_MODBUS.DIP1500_InputRegisters;     // Input registers 0x3001..0x3005
	GVL_COM.COM_DIP1500_1.COM_INPUT_HR_COUNTERS := GVL_MODBUS.DIP1500_Holding_Counters;   // Holding registers 0x4007..0x400A


//------------------------------------------------------------------------------
// HMI : coils (1...)
//------------------------------------------------------------------------------
	//--- DOSENSOR_1
	GVL_COM.COM_DOSENSOR_1.HMI_INPUT_CALIBRATION_HIGH := GVL_MODBUS.Coils_TCP_HMI[0].0;   // 1 | DO Calibration High
	GVL_COM.COM_DOSENSOR_1.HMI_INPUT_CALIBRATION_LOW  := GVL_MODBUS.Coils_TCP_HMI[0].1;   // 2 | DO Calibration Low
	GVL_COM.COM_DOSENSOR_1.HMI_INPUT_LOCAL_REQUEST    := GVL_MODBUS.Coils_TCP_HMI[0].7;   // 8 | DO Sensor Local Request
	GVL_COM.COM_DOSENSOR_1.HMI_INPUT_AUTO_REQUEST     := GVL_MODBUS.Coils_TCP_HMI[1].0;   // 9 | DO Sensor Auto Request

	//--- DIP1500_1
	GVL_COM.COM_DIP1500_1.HMI_INPUT_MOTOR_START_STOP   := GVL_MODBUS.Coils_TCP_HMI[0].2;   // 3 | DIP1500 Motor Start Stop
	GVL_COM.COM_DIP1500_1.HMI_INPUT_MOTOR_DIRECTION    := GVL_MODBUS.Coils_TCP_HMI[0].3;   // 4 | DIP1500 Motor Direction
	GVL_COM.COM_DIP1500_1.HMI_INPUT_FLASH_SAVE         := GVL_MODBUS.Coils_TCP_HMI[0].4;   // 5 | DIP1500 Flash Save
	GVL_COM.COM_DIP1500_1.HMI_INPUT_OPERATION_MODE     := GVL_MODBUS.Coils_TCP_HMI[0].5;   // 6 | DIP1500 Operation Mode
	GVL_COM.COM_DIP1500_1.HMI_INPUT_PARAM_WRITE_ENABLE := GVL_MODBUS.Coils_TCP_HMI[0].6;   // 7 | DIP1500 Parameter Write Enable
	GVL_COM.COM_DIP1500_1.HMI_INPUT_LOCAL_REQUEST      := GVL_MODBUS.Coils_TCP_HMI[1].1;   // 10 | DIP1500 Local Request
	GVL_COM.COM_DIP1500_1.HMI_INPUT_AUTO_REQUEST       := GVL_MODBUS.Coils_TCP_HMI[1].2;   // 11 | DIP1500 Auto Request

	//--- ADM100W_1
	GVL_COM.COM_ADM100W_1.HMI_INPUT_LOCAL_REQUEST := GVL_MODBUS.Coils_TCP_HMI[1].3;   // 12 | ADM100W Local Request
	GVL_COM.COM_ADM100W_1.HMI_INPUT_AUTO_REQUEST  := GVL_MODBUS.Coils_TCP_HMI[1].4;   // 13 | ADM100W Auto Request

	//--- UPI_LOCAL_HMI
	GVL_COM.COM_UPI_LOCAL_HMI.HMI_INPUT_LOCAL_REQUEST := GVL_MODBUS.Coils_TCP_HMI[1].5;   // 14 | Global Local HMI Request
	GVL_COM.COM_UPI_LOCAL_HMI.HMI_INPUT_AUTO_REQUEST  := GVL_MODBUS.Coils_TCP_HMI[1].6;   // 15 | Global Auto HMI Request


//------------------------------------------------------------------------------
// HMI : holding registers (1...), REAL = low word first
//------------------------------------------------------------------------------
	//--- DIP1500_1
	GVL_COM.COM_DIP1500_1.HMI_INPUT_MOTOR_SPEED.Word_value[0]                                := GVL_MODBUS.Holding_register_TCP_HMI[0];   // 1 | DIP1500 Motor Speed (low word)
	GVL_COM.COM_DIP1500_1.HMI_INPUT_MOTOR_SPEED.Word_value[1]                                := GVL_MODBUS.Holding_register_TCP_HMI[1];   // 2 | DIP1500 Motor Speed (high word)
	GVL_COM.COM_DIP1500_1.HMI_INPUT_MAX_MOTOR_SPEED.Word_value[0]                            := GVL_MODBUS.Holding_register_TCP_HMI[2];   // 3 | DIP1500 Max Motor Speed (low word)
	GVL_COM.COM_DIP1500_1.HMI_INPUT_MAX_MOTOR_SPEED.Word_value[1]                            := GVL_MODBUS.Holding_register_TCP_HMI[3];   // 4 | DIP1500 Max Motor Speed (high word)
	GVL_COM.COM_DIP1500_1.HMI_INPUT_RUN_TIME_OR_VOLUME_SETPOINT.Word_value[0]                := GVL_MODBUS.Holding_register_TCP_HMI[4];   // 5 | DIP1500 Run Time Or Volume Setpoint (low word)
	GVL_COM.COM_DIP1500_1.HMI_INPUT_RUN_TIME_OR_VOLUME_SETPOINT.Word_value[1]                := GVL_MODBUS.Holding_register_TCP_HMI[5];   // 6 | DIP1500 Run Time Or Volume Setpoint (high word)
	GVL_COM.COM_DIP1500_1.HMI_INPUT_FLOW_RATE_OR_SPEED_CALIBRATION_COEFFICIENT.Word_value[0] := GVL_MODBUS.Holding_register_TCP_HMI[6];   // 7 | DIP1500 Flow Rate Or Speed Calibration Coefficient (low word)
	GVL_COM.COM_DIP1500_1.HMI_INPUT_FLOW_RATE_OR_SPEED_CALIBRATION_COEFFICIENT.Word_value[1] := GVL_MODBUS.Holding_register_TCP_HMI[7];   // 8 | DIP1500 Flow Rate Or Speed Calibration Coefficient (high word)
	GVL_COM.COM_DIP1500_1.HMI_INPUT_FOOT_SWITCH_INPUT_MODE                                   := GVL_MODBUS.Holding_register_TCP_HMI[8];   // 9 | DIP1500 Foot Switch Input Mode
	GVL_COM.COM_DIP1500_1.HMI_INPUT_LIQUID_LEVEL_INPUT_MODE                                  := GVL_MODBUS.Holding_register_TCP_HMI[9];   // 10 | DIP1500 Liquid Level Input Mode
	GVL_COM.COM_DIP1500_1.HMI_INPUT_STATE_OUTPUT_MODE                                        := GVL_MODBUS.Holding_register_TCP_HMI[10];   // 11 | DIP1500 State Output Mode
	GVL_COM.COM_DIP1500_1.HMI_INPUT_COMMUNICATION_ADDRESS                                    := GVL_MODBUS.Holding_register_TCP_HMI[11];   // 12 | DIP1500 Communication Address
	GVL_COM.COM_DIP1500_1.HMI_INPUT_BAUD_RATE_INDEX                                          := GVL_MODBUS.Holding_register_TCP_HMI[12];   // 13 | DIP1500 Baud Rate Index

GFC_COM_IN := TRUE;

                
END_FUNCTION

FUNCTION GFC_COM_OUT : BOOL

                  
//==============================================================================
// GFC_COM_OUT
// GVL_COM -> Modbus (GVL_MODBUS) : RTU equipment, HMI
// Simple copies only, no conversion (conversions are done in the FBs)
//==============================================================================

//------------------------------------------------------------------------------
// COM : Modbus RTU, to equipment (write triggers are mapped directly in the slave I/O mapping)
//------------------------------------------------------------------------------
	//--- DIP1500_1
	GVL_MODBUS.DIP1500_Coils          := GVL_COM.COM_DIP1500_1.COM_OUTPUT_COILS;       // Coils 0x0001..0x0004
	GVL_MODBUS.DIP1500_Holding_Cmd    := GVL_COM.COM_DIP1500_1.COM_OUTPUT_HR_CMD;      // Holding registers 0x4001..0x4006
	GVL_MODBUS.DIP1500_Holding_Config := GVL_COM.COM_DIP1500_1.COM_OUTPUT_HR_CONFIG;   // Holding registers 0x400B..0x4011


//------------------------------------------------------------------------------
// HMI : discrete inputs (10001...)
//------------------------------------------------------------------------------
	//--- DOSENSOR_1
	GVL_MODBUS.Discret_input_TCP_HMI[0].0 := GVL_COM.COM_DOSENSOR_1.HMI_OUTPUT_FAULT;              // 10001 | Do sensor fault
	GVL_MODBUS.Discret_input_TCP_HMI[0].1 := GVL_COM.COM_DOSENSOR_1.HMI_OUTPUT_CALIBRATION_DONE;   // 10002 | Do sensor calibration done
	GVL_MODBUS.Discret_input_TCP_HMI[1].5 := GVL_COM.COM_DOSENSOR_1.HMI_OUTPUT_LOCAL_ACTIVE;       // 10014 | DO Sensor Local Active

	//--- ADM100W_1
	GVL_MODBUS.Discret_input_TCP_HMI[0].2 := GVL_COM.COM_ADM100W_1.HMI_OUTPUT_ALARM_1_STATUS;    // 10003 | ADM100W Alarm 1 Status
	GVL_MODBUS.Discret_input_TCP_HMI[0].3 := GVL_COM.COM_ADM100W_1.HMI_OUTPUT_ALARM_2_STATUS;    // 10004 | ADM100W Alarm 2 Status
	GVL_MODBUS.Discret_input_TCP_HMI[0].4 := GVL_COM.COM_ADM100W_1.HMI_OUTPUT_ALARM_3_STATUS;    // 10005 | ADM100W Alarm 3 Status
	GVL_MODBUS.Discret_input_TCP_HMI[0].5 := GVL_COM.COM_ADM100W_1.HMI_OUTPUT_ALARM_4_STATUS;    // 10006 | ADM100W Alarm 4 Status
	GVL_MODBUS.Discret_input_TCP_HMI[0].6 := GVL_COM.COM_ADM100W_1.HMI_OUTPUT_ALARM_5_STATUS;    // 10007 | ADM100W Alarm 5 Status
	GVL_MODBUS.Discret_input_TCP_HMI[0].7 := GVL_COM.COM_ADM100W_1.HMI_OUTPUT_ALARM_6_STATUS;    // 10008 | ADM100W Alarm 6 Status
	GVL_MODBUS.Discret_input_TCP_HMI[1].0 := GVL_COM.COM_ADM100W_1.HMI_OUTPUT_ALARM_7_STATUS;    // 10009 | ADM100W Alarm 7 Status
	GVL_MODBUS.Discret_input_TCP_HMI[1].1 := GVL_COM.COM_ADM100W_1.HMI_OUTPUT_ALARM_8_STATUS;    // 10010 | ADM100W Alarm 8 Status
	GVL_MODBUS.Discret_input_TCP_HMI[1].2 := GVL_COM.COM_ADM100W_1.HMI_OUTPUT_ALARM_9_STATUS;    // 10011 | ADM100W Alarm 9 Status
	GVL_MODBUS.Discret_input_TCP_HMI[1].3 := GVL_COM.COM_ADM100W_1.HMI_OUTPUT_ALARM_10_STATUS;   // 10012 | ADM100W Alarm 10 Status
	GVL_MODBUS.Discret_input_TCP_HMI[2].1 := GVL_COM.COM_ADM100W_1.HMI_OUTPUT_LOCAL_ACTIVE;      // 10018 | ADM100W Local Active

	//--- DIP1500_1
	GVL_MODBUS.Discret_input_TCP_HMI[1].7 := GVL_COM.COM_DIP1500_1.HMI_OUTPUT_LOCAL_ACTIVE;   // 10016 | DIP1500 Local Active

	//--- UPI_LOCAL_HMI
	GVL_MODBUS.Discret_input_TCP_HMI[2].3 := GVL_COM.COM_UPI_LOCAL_HMI.HMI_OUTPUT_LOCAL_ACTIVE;   // 10020 | Global Local HMI Active


//------------------------------------------------------------------------------
// HMI : input registers (1...), REAL = low word first
//------------------------------------------------------------------------------
	//--- ADM100W_1
	GVL_MODBUS.Input_register_TCP_HMI[0] := GVL_COM.COM_ADM100W_1.HMI_OUTPUT_FREQUENCY.Word_value[0];                   // 1 | ADM100W Frequency (low word)
	GVL_MODBUS.Input_register_TCP_HMI[1] := GVL_COM.COM_ADM100W_1.HMI_OUTPUT_FREQUENCY.Word_value[1];                   // 2 | ADM100W Frequency (high word)
	GVL_MODBUS.Input_register_TCP_HMI[2] := GVL_COM.COM_ADM100W_1.HMI_OUTPUT_L1_L2_VOLTAGE.Word_value[0];               // 3 | ADM100W L1-L2 Voltage (low word)
	GVL_MODBUS.Input_register_TCP_HMI[3] := GVL_COM.COM_ADM100W_1.HMI_OUTPUT_L1_L2_VOLTAGE.Word_value[1];               // 4 | ADM100W L1-L2 Voltage (high word)
	GVL_MODBUS.Input_register_TCP_HMI[4] := GVL_COM.COM_ADM100W_1.HMI_OUTPUT_L1_N_VOLTAGE.Word_value[0];                // 5 | ADM100W L1-N Voltage (low word)
	GVL_MODBUS.Input_register_TCP_HMI[5] := GVL_COM.COM_ADM100W_1.HMI_OUTPUT_L1_N_VOLTAGE.Word_value[1];                // 6 | ADM100W L1-N Voltage (high word)
	GVL_MODBUS.Input_register_TCP_HMI[6] := GVL_COM.COM_ADM100W_1.HMI_OUTPUT_L1_CURRENT.Word_value[0];                  // 7 | ADM100W L1 Current (low word)
	GVL_MODBUS.Input_register_TCP_HMI[7] := GVL_COM.COM_ADM100W_1.HMI_OUTPUT_L1_CURRENT.Word_value[1];                  // 8 | ADM100W L1 Current (high word)
	GVL_MODBUS.Input_register_TCP_HMI[8] := GVL_COM.COM_ADM100W_1.HMI_OUTPUT_L1_ACTIVE_POWER.Word_value[0];             // 9 | ADM100W L1 Active Power (low word)
	GVL_MODBUS.Input_register_TCP_HMI[9] := GVL_COM.COM_ADM100W_1.HMI_OUTPUT_L1_ACTIVE_POWER.Word_value[1];             // 10 | ADM100W L1 Active Power (high word)
	GVL_MODBUS.Input_register_TCP_HMI[10] := GVL_COM.COM_ADM100W_1.HMI_OUTPUT_L1_APPARENT_POWER.Word_value[0];           // 11 | ADM100W L1 Apparent Power (low word)
	GVL_MODBUS.Input_register_TCP_HMI[11] := GVL_COM.COM_ADM100W_1.HMI_OUTPUT_L1_APPARENT_POWER.Word_value[1];           // 12 | ADM100W L1 Apparent Power (high word)
	GVL_MODBUS.Input_register_TCP_HMI[12] := GVL_COM.COM_ADM100W_1.HMI_OUTPUT_L1_REACTIVE_POWER.Word_value[0];           // 13 | ADM100W L1 Reactive Power (low word)
	GVL_MODBUS.Input_register_TCP_HMI[13] := GVL_COM.COM_ADM100W_1.HMI_OUTPUT_L1_REACTIVE_POWER.Word_value[1];           // 14 | ADM100W L1 Reactive Power (high word)
	GVL_MODBUS.Input_register_TCP_HMI[14] := GVL_COM.COM_ADM100W_1.HMI_OUTPUT_L1_CURRENT_PHASE_ANGLE.Word_value[0];      // 15 | ADM100W L1 Current Phase Angle (low word)
	GVL_MODBUS.Input_register_TCP_HMI[15] := GVL_COM.COM_ADM100W_1.HMI_OUTPUT_L1_CURRENT_PHASE_ANGLE.Word_value[1];      // 16 | ADM100W L1 Current Phase Angle (high word)
	GVL_MODBUS.Input_register_TCP_HMI[16] := GVL_COM.COM_ADM100W_1.HMI_OUTPUT_L1_POWER_FACTOR.Word_value[0];             // 17 | ADM100W L1 Power Factor (low word)
	GVL_MODBUS.Input_register_TCP_HMI[17] := GVL_COM.COM_ADM100W_1.HMI_OUTPUT_L1_POWER_FACTOR.Word_value[1];             // 18 | ADM100W L1 Power Factor (high word)
	GVL_MODBUS.Input_register_TCP_HMI[18] := GVL_COM.COM_ADM100W_1.HMI_OUTPUT_L1_VOLTAGE_THD.Word_value[0];              // 19 | ADM100W L1 Voltage THD (low word)
	GVL_MODBUS.Input_register_TCP_HMI[19] := GVL_COM.COM_ADM100W_1.HMI_OUTPUT_L1_VOLTAGE_THD.Word_value[1];              // 20 | ADM100W L1 Voltage THD (high word)
	GVL_MODBUS.Input_register_TCP_HMI[20] := GVL_COM.COM_ADM100W_1.HMI_OUTPUT_L1_CURRENT_THD.Word_value[0];              // 21 | ADM100W L1 Current THD (low word)
	GVL_MODBUS.Input_register_TCP_HMI[21] := GVL_COM.COM_ADM100W_1.HMI_OUTPUT_L1_CURRENT_THD.Word_value[1];              // 22 | ADM100W L1 Current THD (high word)
	GVL_MODBUS.Input_register_TCP_HMI[22] := GVL_COM.COM_ADM100W_1.HMI_OUTPUT_L1_MAX_LOAD.Word_value[0];                 // 23 | ADM100W L1 Max Load (low word)
	GVL_MODBUS.Input_register_TCP_HMI[23] := GVL_COM.COM_ADM100W_1.HMI_OUTPUT_L1_MAX_LOAD.Word_value[1];                 // 24 | ADM100W L1 Max Load (high word)
	GVL_MODBUS.Input_register_TCP_HMI[24] := GVL_COM.COM_ADM100W_1.HMI_OUTPUT_L1_L2_VOLTAGE_PHASE_ANGLE.Word_value[0];   // 25 | ADM100W L1-L2 Voltage Phase Angle (low word)
	GVL_MODBUS.Input_register_TCP_HMI[25] := GVL_COM.COM_ADM100W_1.HMI_OUTPUT_L1_L2_VOLTAGE_PHASE_ANGLE.Word_value[1];   // 26 | ADM100W L1-L2 Voltage Phase Angle (high word)
	GVL_MODBUS.Input_register_TCP_HMI[26] := GVL_COM.COM_ADM100W_1.HMI_OUTPUT_L2_L3_VOLTAGE.Word_value[0];               // 27 | ADM100W L2-L3 Voltage (low word)
	GVL_MODBUS.Input_register_TCP_HMI[27] := GVL_COM.COM_ADM100W_1.HMI_OUTPUT_L2_L3_VOLTAGE.Word_value[1];               // 28 | ADM100W L2-L3 Voltage (high word)
	GVL_MODBUS.Input_register_TCP_HMI[28] := GVL_COM.COM_ADM100W_1.HMI_OUTPUT_L2_N_VOLTAGE.Word_value[0];                // 29 | ADM100W L2-N Voltage (low word)
	GVL_MODBUS.Input_register_TCP_HMI[29] := GVL_COM.COM_ADM100W_1.HMI_OUTPUT_L2_N_VOLTAGE.Word_value[1];                // 30 | ADM100W L2-N Voltage (high word)
	GVL_MODBUS.Input_register_TCP_HMI[30] := GVL_COM.COM_ADM100W_1.HMI_OUTPUT_L2_CURRENT.Word_value[0];                  // 31 | ADM100W L2 Current (low word)
	GVL_MODBUS.Input_register_TCP_HMI[31] := GVL_COM.COM_ADM100W_1.HMI_OUTPUT_L2_CURRENT.Word_value[1];                  // 32 | ADM100W L2 Current (high word)
	GVL_MODBUS.Input_register_TCP_HMI[32] := GVL_COM.COM_ADM100W_1.HMI_OUTPUT_L2_ACTIVE_POWER.Word_value[0];             // 33 | ADM100W L2 Active Power (low word)
	GVL_MODBUS.Input_register_TCP_HMI[33] := GVL_COM.COM_ADM100W_1.HMI_OUTPUT_L2_ACTIVE_POWER.Word_value[1];             // 34 | ADM100W L2 Active Power (high word)
	GVL_MODBUS.Input_register_TCP_HMI[34] := GVL_COM.COM_ADM100W_1.HMI_OUTPUT_L2_APPARENT_POWER.Word_value[0];           // 35 | ADM100W L2 Apparent Power (low word)
	GVL_MODBUS.Input_register_TCP_HMI[35] := GVL_COM.COM_ADM100W_1.HMI_OUTPUT_L2_APPARENT_POWER.Word_value[1];           // 36 | ADM100W L2 Apparent Power (high word)
	GVL_MODBUS.Input_register_TCP_HMI[36] := GVL_COM.COM_ADM100W_1.HMI_OUTPUT_L2_REACTIVE_POWER.Word_value[0];           // 37 | ADM100W L2 Reactive Power (low word)
	GVL_MODBUS.Input_register_TCP_HMI[37] := GVL_COM.COM_ADM100W_1.HMI_OUTPUT_L2_REACTIVE_POWER.Word_value[1];           // 38 | ADM100W L2 Reactive Power (high word)
	GVL_MODBUS.Input_register_TCP_HMI[38] := GVL_COM.COM_ADM100W_1.HMI_OUTPUT_L2_CURRENT_PHASE_ANGLE.Word_value[0];      // 39 | ADM100W L2 Current Phase Angle (low word)
	GVL_MODBUS.Input_register_TCP_HMI[39] := GVL_COM.COM_ADM100W_1.HMI_OUTPUT_L2_CURRENT_PHASE_ANGLE.Word_value[1];      // 40 | ADM100W L2 Current Phase Angle (high word)
	GVL_MODBUS.Input_register_TCP_HMI[40] := GVL_COM.COM_ADM100W_1.HMI_OUTPUT_L2_POWER_FACTOR.Word_value[0];             // 41 | ADM100W L2 Power Factor (low word)
	GVL_MODBUS.Input_register_TCP_HMI[41] := GVL_COM.COM_ADM100W_1.HMI_OUTPUT_L2_POWER_FACTOR.Word_value[1];             // 42 | ADM100W L2 Power Factor (high word)
	GVL_MODBUS.Input_register_TCP_HMI[42] := GVL_COM.COM_ADM100W_1.HMI_OUTPUT_L2_VOLTAGE_THD.Word_value[0];              // 43 | ADM100W L2 Voltage THD (low word)
	GVL_MODBUS.Input_register_TCP_HMI[43] := GVL_COM.COM_ADM100W_1.HMI_OUTPUT_L2_VOLTAGE_THD.Word_value[1];              // 44 | ADM100W L2 Voltage THD (high word)
	GVL_MODBUS.Input_register_TCP_HMI[44] := GVL_COM.COM_ADM100W_1.HMI_OUTPUT_L2_CURRENT_THD.Word_value[0];              // 45 | ADM100W L2 Current THD (low word)
	GVL_MODBUS.Input_register_TCP_HMI[45] := GVL_COM.COM_ADM100W_1.HMI_OUTPUT_L2_CURRENT_THD.Word_value[1];              // 46 | ADM100W L2 Current THD (high word)
	GVL_MODBUS.Input_register_TCP_HMI[46] := GVL_COM.COM_ADM100W_1.HMI_OUTPUT_L2_MAX_LOAD.Word_value[0];                 // 47 | ADM100W L2 Max Load (low word)
	GVL_MODBUS.Input_register_TCP_HMI[47] := GVL_COM.COM_ADM100W_1.HMI_OUTPUT_L2_MAX_LOAD.Word_value[1];                 // 48 | ADM100W L2 Max Load (high word)
	GVL_MODBUS.Input_register_TCP_HMI[48] := GVL_COM.COM_ADM100W_1.HMI_OUTPUT_L1_L3_VOLTAGE_PHASE_ANGLE.Word_value[0];   // 49 | ADM100W L1-L3 Voltage Phase Angle (low word)
	GVL_MODBUS.Input_register_TCP_HMI[49] := GVL_COM.COM_ADM100W_1.HMI_OUTPUT_L1_L3_VOLTAGE_PHASE_ANGLE.Word_value[1];   // 50 | ADM100W L1-L3 Voltage Phase Angle (high word)
	GVL_MODBUS.Input_register_TCP_HMI[50] := GVL_COM.COM_ADM100W_1.HMI_OUTPUT_L3_L1_VOLTAGE.Word_value[0];               // 51 | ADM100W L3-L1 Voltage (low word)
	GVL_MODBUS.Input_register_TCP_HMI[51] := GVL_COM.COM_ADM100W_1.HMI_OUTPUT_L3_L1_VOLTAGE.Word_value[1];               // 52 | ADM100W L3-L1 Voltage (high word)
	GVL_MODBUS.Input_register_TCP_HMI[52] := GVL_COM.COM_ADM100W_1.HMI_OUTPUT_L3_N_VOLTAGE.Word_value[0];                // 53 | ADM100W L3-N Voltage (low word)
	GVL_MODBUS.Input_register_TCP_HMI[53] := GVL_COM.COM_ADM100W_1.HMI_OUTPUT_L3_N_VOLTAGE.Word_value[1];                // 54 | ADM100W L3-N Voltage (high word)
	GVL_MODBUS.Input_register_TCP_HMI[54] := GVL_COM.COM_ADM100W_1.HMI_OUTPUT_L3_CURRENT.Word_value[0];                  // 55 | ADM100W L3 Current (low word)
	GVL_MODBUS.Input_register_TCP_HMI[55] := GVL_COM.COM_ADM100W_1.HMI_OUTPUT_L3_CURRENT.Word_value[1];                  // 56 | ADM100W L3 Current (high word)
	GVL_MODBUS.Input_register_TCP_HMI[56] := GVL_COM.COM_ADM100W_1.HMI_OUTPUT_L3_ACTIVE_POWER.Word_value[0];             // 57 | ADM100W L3 Active Power (low word)
	GVL_MODBUS.Input_register_TCP_HMI[57] := GVL_COM.COM_ADM100W_1.HMI_OUTPUT_L3_ACTIVE_POWER.Word_value[1];             // 58 | ADM100W L3 Active Power (high word)
	GVL_MODBUS.Input_register_TCP_HMI[58] := GVL_COM.COM_ADM100W_1.HMI_OUTPUT_L3_APPARENT_POWER.Word_value[0];           // 59 | ADM100W L3 Apparent Power (low word)
	GVL_MODBUS.Input_register_TCP_HMI[59] := GVL_COM.COM_ADM100W_1.HMI_OUTPUT_L3_APPARENT_POWER.Word_value[1];           // 60 | ADM100W L3 Apparent Power (high word)
	GVL_MODBUS.Input_register_TCP_HMI[60] := GVL_COM.COM_ADM100W_1.HMI_OUTPUT_L3_REACTIVE_POWER.Word_value[0];           // 61 | ADM100W L3 Reactive Power (low word)
	GVL_MODBUS.Input_register_TCP_HMI[61] := GVL_COM.COM_ADM100W_1.HMI_OUTPUT_L3_REACTIVE_POWER.Word_value[1];           // 62 | ADM100W L3 Reactive Power (high word)
	GVL_MODBUS.Input_register_TCP_HMI[62] := GVL_COM.COM_ADM100W_1.HMI_OUTPUT_L3_CURRENT_PHASE_ANGLE.Word_value[0];      // 63 | ADM100W L3 Current Phase Angle (low word)
	GVL_MODBUS.Input_register_TCP_HMI[63] := GVL_COM.COM_ADM100W_1.HMI_OUTPUT_L3_CURRENT_PHASE_ANGLE.Word_value[1];      // 64 | ADM100W L3 Current Phase Angle (high word)
	GVL_MODBUS.Input_register_TCP_HMI[64] := GVL_COM.COM_ADM100W_1.HMI_OUTPUT_L3_POWER_FACTOR.Word_value[0];             // 65 | ADM100W L3 Power Factor (low word)
	GVL_MODBUS.Input_register_TCP_HMI[65] := GVL_COM.COM_ADM100W_1.HMI_OUTPUT_L3_POWER_FACTOR.Word_value[1];             // 66 | ADM100W L3 Power Factor (high word)
	GVL_MODBUS.Input_register_TCP_HMI[66] := GVL_COM.COM_ADM100W_1.HMI_OUTPUT_L3_VOLTAGE_THD.Word_value[0];              // 67 | ADM100W L3 Voltage THD (low word)
	GVL_MODBUS.Input_register_TCP_HMI[67] := GVL_COM.COM_ADM100W_1.HMI_OUTPUT_L3_VOLTAGE_THD.Word_value[1];              // 68 | ADM100W L3 Voltage THD (high word)
	GVL_MODBUS.Input_register_TCP_HMI[68] := GVL_COM.COM_ADM100W_1.HMI_OUTPUT_L3_CURRENT_THD.Word_value[0];              // 69 | ADM100W L3 Current THD (low word)
	GVL_MODBUS.Input_register_TCP_HMI[69] := GVL_COM.COM_ADM100W_1.HMI_OUTPUT_L3_CURRENT_THD.Word_value[1];              // 70 | ADM100W L3 Current THD (high word)
	GVL_MODBUS.Input_register_TCP_HMI[70] := GVL_COM.COM_ADM100W_1.HMI_OUTPUT_L3_MAX_LOAD.Word_value[0];                 // 71 | ADM100W L3 Max Load (low word)
	GVL_MODBUS.Input_register_TCP_HMI[71] := GVL_COM.COM_ADM100W_1.HMI_OUTPUT_L3_MAX_LOAD.Word_value[1];                 // 72 | ADM100W L3 Max Load (high word)
	GVL_MODBUS.Input_register_TCP_HMI[72] := GVL_COM.COM_ADM100W_1.HMI_OUTPUT_INTERNAL_TEMPERATURE.Word_value[0];        // 73 | ADM100W Internal Temperature (low word)
	GVL_MODBUS.Input_register_TCP_HMI[73] := GVL_COM.COM_ADM100W_1.HMI_OUTPUT_INTERNAL_TEMPERATURE.Word_value[1];        // 74 | ADM100W Internal Temperature (high word)
	GVL_MODBUS.Input_register_TCP_HMI[74] := GVL_COM.COM_ADM100W_1.HMI_OUTPUT_ACTIVE_ENERGY.Word_value[0];               // 75 | ADM100W Active Energy (low word)
	GVL_MODBUS.Input_register_TCP_HMI[75] := GVL_COM.COM_ADM100W_1.HMI_OUTPUT_ACTIVE_ENERGY.Word_value[1];               // 76 | ADM100W Active Energy (high word)
	GVL_MODBUS.Input_register_TCP_HMI[76] := GVL_COM.COM_ADM100W_1.HMI_OUTPUT_APPARENT_ENERGY.Word_value[0];             // 77 | ADM100W Apparent Energy (low word)
	GVL_MODBUS.Input_register_TCP_HMI[77] := GVL_COM.COM_ADM100W_1.HMI_OUTPUT_APPARENT_ENERGY.Word_value[1];             // 78 | ADM100W Apparent Energy (high word)
	GVL_MODBUS.Input_register_TCP_HMI[78] := GVL_COM.COM_ADM100W_1.HMI_OUTPUT_REACTIVE_ENERGY.Word_value[0];             // 79 | ADM100W Reactive Energy (low word)
	GVL_MODBUS.Input_register_TCP_HMI[79] := GVL_COM.COM_ADM100W_1.HMI_OUTPUT_REACTIVE_ENERGY.Word_value[1];             // 80 | ADM100W Reactive Energy (high word)
	GVL_MODBUS.Input_register_TCP_HMI[80] := GVL_COM.COM_ADM100W_1.HMI_OUTPUT_TOTAL_ACTIVE_POWER.Word_value[0];          // 81 | ADM100W Total Active Power (low word)
	GVL_MODBUS.Input_register_TCP_HMI[81] := GVL_COM.COM_ADM100W_1.HMI_OUTPUT_TOTAL_ACTIVE_POWER.Word_value[1];          // 82 | ADM100W Total Active Power (high word)
	GVL_MODBUS.Input_register_TCP_HMI[82] := GVL_COM.COM_ADM100W_1.HMI_OUTPUT_TOTAL_APPARENT_POWER.Word_value[0];        // 83 | ADM100W Total Apparent Power (low word)
	GVL_MODBUS.Input_register_TCP_HMI[83] := GVL_COM.COM_ADM100W_1.HMI_OUTPUT_TOTAL_APPARENT_POWER.Word_value[1];        // 84 | ADM100W Total Apparent Power (high word)
	GVL_MODBUS.Input_register_TCP_HMI[84] := GVL_COM.COM_ADM100W_1.HMI_OUTPUT_TOTAL_REACTIVE_POWER.Word_value[0];        // 85 | ADM100W Total Reactive Power (low word)
	GVL_MODBUS.Input_register_TCP_HMI[85] := GVL_COM.COM_ADM100W_1.HMI_OUTPUT_TOTAL_REACTIVE_POWER.Word_value[1];        // 86 | ADM100W Total Reactive Power (high word)
	GVL_MODBUS.Input_register_TCP_HMI[86] := GVL_COM.COM_ADM100W_1.HMI_OUTPUT_ALL_PHASE_POWER_FACTOR.Word_value[0];      // 87 | ADM100W All Phase Power Factor (low word)
	GVL_MODBUS.Input_register_TCP_HMI[87] := GVL_COM.COM_ADM100W_1.HMI_OUTPUT_ALL_PHASE_POWER_FACTOR.Word_value[1];      // 88 | ADM100W All Phase Power Factor (high word)

	//--- DOSENSOR_1
	GVL_MODBUS.Input_register_TCP_HMI[88] := GVL_COM.COM_DOSENSOR_1.HMI_OUTPUT_SIGNAL.Word_value[0];   // 89 | DO Sensor Signal (low word)
	GVL_MODBUS.Input_register_TCP_HMI[89] := GVL_COM.COM_DOSENSOR_1.HMI_OUTPUT_SIGNAL.Word_value[1];   // 90 | DO Sensor Signal (high word)

	//--- DIP1500_1
	GVL_MODBUS.Input_register_TCP_HMI[90] := GVL_COM.COM_DIP1500_1.HMI_OUTPUT_FIRMWARE_VERSION;                               // 91 | DIP1500 Firmware Version
	GVL_MODBUS.Input_register_TCP_HMI[91] := GVL_COM.COM_DIP1500_1.HMI_OUTPUT_HARDWARE_VERSION;                               // 92 | DIP1500 Hardware Version
	GVL_MODBUS.Input_register_TCP_HMI[92] := GVL_COM.COM_DIP1500_1.HMI_OUTPUT_TEMPERATURE;                                    // 93 | DIP1500 Temperature
	GVL_MODBUS.Input_register_TCP_HMI[93] := GVL_COM.COM_DIP1500_1.HMI_OUTPUT_FLOAT_LEVEL_ALARM;                              // 94 | DIP1500 Float Level Alarm
	GVL_MODBUS.Input_register_TCP_HMI[94] := GVL_COM.COM_DIP1500_1.HMI_OUTPUT_DIGITAL_OUTPUT_VALUE;                           // 95 | DIP1500 Digital Output Value
	GVL_MODBUS.Input_register_TCP_HMI[95] := GVL_COM.COM_DIP1500_1.HMI_OUTPUT_REAL_TIME_RUN_TIME_OR_VOLUME.Word_value[0];     // 96 | DIP1500 Real-Time Run Time Or Volume (low word)
	GVL_MODBUS.Input_register_TCP_HMI[96] := GVL_COM.COM_DIP1500_1.HMI_OUTPUT_REAL_TIME_RUN_TIME_OR_VOLUME.Word_value[1];     // 97 | DIP1500 Real-Time Run Time Or Volume (high word)
	GVL_MODBUS.Input_register_TCP_HMI[97] := GVL_COM.COM_DIP1500_1.HMI_OUTPUT_ACCUMULATED_RUN_TIME_OR_VOLUME.Word_value[0];   // 98 | DIP1500 Accumulated Run Time Or Volume (low word)
	GVL_MODBUS.Input_register_TCP_HMI[98] := GVL_COM.COM_DIP1500_1.HMI_OUTPUT_ACCUMULATED_RUN_TIME_OR_VOLUME.Word_value[1];   // 99 | DIP1500 Accumulated Run Time Or Volume (high word)

GFC_COM_OUT := TRUE;

                
END_FUNCTION

FUNCTION GFC_EXC : BOOL

                  
//==============================================================================
// GFC_EXC
// Exchanges between instances : one FC_EXC_<A>_<B> call per pair of instances
// Called after GFB_UPI and before GFB_INST
//==============================================================================

//------------------------------------------------------------------------------
// ADM100W_1
//------------------------------------------------------------------------------
	//--- UPI_LOCAL_HMI <-> ADM100W_1
	FC_EXC_UPI_LOCAL_HMI_ADM100W(
		EXC_UPI_LOCAL_HMI := GVL_EXC.EXC_UPI_LOCAL_HMI,
		EXC_ADM100W       := GVL_EXC.EXC_ADM100W_1);


//------------------------------------------------------------------------------
// DOSENSOR_1
//------------------------------------------------------------------------------
	//--- UPI_LOCAL_HMI <-> DOSENSOR_1
	FC_EXC_UPI_LOCAL_HMI_DOSENSOR(
		EXC_UPI_LOCAL_HMI := GVL_EXC.EXC_UPI_LOCAL_HMI,
		EXC_DOSENSOR      := GVL_EXC.EXC_DOSENSOR_1);


//------------------------------------------------------------------------------
// DIP1500_1
//------------------------------------------------------------------------------
	//--- UPI_LOCAL_HMI <-> DIP1500_1
	FC_EXC_UPI_LOCAL_HMI_DIP1500(
		EXC_UPI_LOCAL_HMI := GVL_EXC.EXC_UPI_LOCAL_HMI,
		EXC_DIP1500       := GVL_EXC.EXC_DIP1500_1);

GFC_EXC := TRUE;

                
END_FUNCTION

FUNCTION GFC_IO_IN : BOOL

                  
//==============================================================================
// GFC_IO_IN
// GVL_IOMAP (PLC I/O cards) -> GVL_IO
// Simple copies only, no conversion (conversions are done in the FBs)
//==============================================================================

//------------------------------------------------------------------------------
// Digital inputs
//------------------------------------------------------------------------------
	//--- DOSENSOR_1
	GVL_IO.IO_DOSENSOR_1.INPUT_SENSOR_FAULT := GVL_IOMAP.IOMAP_DI_FAULT_DOSENSOR_1;


//------------------------------------------------------------------------------
// Analog inputs
//------------------------------------------------------------------------------
	//--- DOSENSOR_1
	GVL_IO.IO_DOSENSOR_1.INPUT_SIGNAL := GVL_IOMAP.IOMAP_AI_SIGNAL_DOSENSOR_1;

GFC_IO_IN := TRUE;

                
END_FUNCTION

FUNCTION GFC_IO_OUT : BOOL

                  
//==============================================================================
// GFC_IO_OUT
// GVL_IO -> GVL_IOMAP (PLC I/O cards)
// Simple copies only, no conversion (conversions are done in the FBs)
//==============================================================================

//------------------------------------------------------------------------------
// Digital outputs
//------------------------------------------------------------------------------
	//--- DOSENSOR_1
	GVL_IOMAP.IOMAP_DO_HIGH_DOSENSOR_1 := GVL_IO.IO_DOSENSOR_1.OUTPUT_CALIBRATION_HIGH;
	GVL_IOMAP.IOMAP_DO_LOW_DOSENSOR_1  := GVL_IO.IO_DOSENSOR_1.OUTPUT_CALIBRATION_LOW;

GFC_IO_OUT := TRUE;

                
END_FUNCTION

PROGRAM PLC_PRG
  VAR
    GFB_UPI_1 : GFB_UPI;  (* Functional units *)
    GFB_INST_1 : GFB_INST;  (* Equipment instances *)
  END_VAR

                  
//==============================================================================
// PLC_PRG
// Main cycle : 1. read all inputs, 2. functional units, 3. equipment, 4. write all outputs
//==============================================================================

//------------------------------------------------------------------------------
// 1. INPUTS : interfaces -> GVL
//------------------------------------------------------------------------------
GFC_COM_IN();
GFC_IO_IN();

//------------------------------------------------------------------------------
// 2. FUNCTIONAL UNITS (UPI) and exchanges between instances
//------------------------------------------------------------------------------
GFB_UPI_1();
GFC_EXC();      // exchanges between instances (FC_EXC_...)

//------------------------------------------------------------------------------
// 3. EQUIPMENT
//------------------------------------------------------------------------------
GFB_INST_1();

//------------------------------------------------------------------------------
// 4. OUTPUTS : GVL -> interfaces
//------------------------------------------------------------------------------
GFC_COM_OUT();
GFC_IO_OUT();

                
END_PROGRAM

CONFIGURATION Application
  RESOURCE Application ON PLC
    VAR_GLOBAL  (* GVL_MODBUS *)
      Coils_TCP_HMI : ARRAY[0..187] OF BYTE;  (* -----------------Modbus TCP line IHM -> API (coils, %IX) *)
      Discret_input_TCP_HMI : ARRAY[0..187] OF BYTE;  (* API -> IHM (entrées discrètes, %QX) *)
      Holding_register_TCP_HMI : ARRAY[0..1500] OF WORD;  (* IHM -> API (registres de retenue, %IW) *)
      Input_register_TCP_HMI : ARRAY[0..1500] OF WORD;  (* API -> IHM (registres d'entrée, %QW) *)
      ADM100W_InputRegisters : ARRAY[0..87] OF WORD;  (* ------------------Modbus RTU line ---ADM100W *)
      ADM100W_Alarms : ARRAY[0..1] OF BYTE;
      DIP1500_Coils : ARRAY[0..3] OF BOOL;  (* ---Kamoer DIP1500 Coils - wrinting to pump *)
      DIP1500_InputRegisters : ARRAY[0..4] OF WORD;  (* input register - reading from pump *)
      DIP1500_Holding_Cmd : ARRAY[0..5] OF WORD;  (* Discrete input Holding registers - Writing to pump *)
      DIP1500_Holding_Config : ARRAY[0..6] OF WORD;
      DIP1500_Holding_Counters : ARRAY[0..3] OF WORD;  (* Holding registers - Reading from pump *)
    END_VAR
    {attribute 'qualified_only'}
    VAR_GLOBAL  (* GVL_IOMAP *)
      IOMAP_AI_SIGNAL_DOSENSOR_1 : DWORD;
      IOMAP_DI_FAULT_DOSENSOR_1 : BOOL;
      IOMAP_DO_HIGH_DOSENSOR_1 : BOOL;
      IOMAP_DO_LOW_DOSENSOR_1 : BOOL;
    END_VAR
    {attribute 'qualified_only'}
    {attribute 'checksumnoinit_override' := '3446479488'}
    {attribute 'init_related_code' := '6eea8fa9-da21-468e-bab1-ddc04c20a5e9'}
    VAR_GLOBAL RETAIN PERSISTENT  (* GVL_PA *)
      {attribute 'order_in_persistent_editor' := '0'}
      PA_ADM100W_1 : DUT_PA_ADM100W;  (* Trumeter ADM100W power meter *)
      {attribute 'order_in_persistent_editor' := '1'}
      PA_DOSENSOR_1 : DUT_PA_DOSENSOR;  (* Dissolved oxygen sensor *)
      {attribute 'order_in_persistent_editor' := '2'}
      PA_DIP1500_1 : DUT_PA_DIP1500;  (* Kamoer DIP1500 peristaltic pump *)
    END_VAR
    {attribute 'qualified_only'}
    VAR_GLOBAL  (* GVL_COM *)
      COM_ADM100W_1 : DUT_COM_ADM100W;  (* Trumeter ADM100W power meter *)
      COM_DOSENSOR_1 : DUT_COM_DOSENSOR;  (* Dissolved oxygen sensor *)
      COM_DIP1500_1 : DUT_COM_DIP1500;  (* Kamoer DIP1500 peristaltic pump *)
      COM_UPI_LOCAL_HMI : DUT_COM_UPI_LOCAL_HMI;  (* Global HMI local mode *)
    END_VAR
    {attribute 'qualified_only'}
    VAR_GLOBAL  (* GVL_EXC *)
      EXC_ADM100W_1 : DUT_EXC_ADM100W;  (* Trumeter ADM100W power meter *)
      EXC_DOSENSOR_1 : DUT_EXC_DOSENSOR;  (* Dissolved oxygen sensor *)
      EXC_DIP1500_1 : DUT_EXC_DIP1500;  (* Kamoer DIP1500 peristaltic pump *)
      EXC_UPI_LOCAL_HMI : DUT_EXC_UPI_LOCAL_HMI;  (* Global HMI local mode *)
    END_VAR
    {attribute 'qualified_only'}
    VAR_GLOBAL  (* GVL_IO *)
      IO_ADM100W_1 : DUT_IO_ADM100W;  (* Trumeter ADM100W power meter *)
      IO_DOSENSOR_1 : DUT_IO_DOSENSOR;  (* Dissolved oxygen sensor *)
      IO_DIP1500_1 : DUT_IO_DIP1500;  (* Kamoer DIP1500 peristaltic pump *)
    END_VAR
  END_RESOURCE
END_CONFIGURATION
